(* IEC 61131-3 sources: daoli-st-library/DL_Base (part 16) *)

(* ---- FB_DL_SchmittTriggerGap.st ---- *)
(*
  Name        : FB_DL_SchmittTriggerGap
  Category    : DL_Base
  Version     : 1.0.0
  Purpose     : 带回差的双阈值整形器（施密特）：上阈置位、下阈复位，滞带宽可组态，输出干净布尔电平与单拍沿脉冲；/ Dual-threshold Schmitt shaping: set at upper threshold, reset at lower threshold, configurable hysteresis band, clean boolean plus single-scan edge pulses
  溯源        : 借 t2-1-lgf·comparator 的分类/参数域组织，clean-room 实现
  Boundary    : ① 组态闸：fThHigh - fThLow <= eps（带宽容差比较，禁 = ）→ 锁存故障，输出保持 FALSE；
                ② 非有限输入该拍不参与翻转判定（保留上拍电平，防误翻）；
                ③ 翻转计数 UDINT 饱和：到 4294967295 前停止累加（防回绕）；
                ④ 沿脉冲单拍化：内部 _b* 置位 → 出口统一映射，不在 CASE 内直接写输出（R187）。
*)
TYPE E_DL_SchState :
(
    eIdle  := 0,                             (* 未使能 / Disabled *)
    eRun   := 10,                            (* 整形运行 / Shaping active *)
    eFault := 90                             (* 故障锁存相 / Fault latched *)
);
END_TYPE

TYPE E_DL_SchCause :
(
    eNone       := 0,                        (* 无故障成因 / No cause *)
    eCfgIllegal := 1,                        (* 组态非法：滞带宽非正 / Illegal config: band non-positive *)
    ePhaseBad   := 2                         (* 非法相位兜底 / Illegal phase fallback *)
);
END_TYPE

FUNCTION_BLOCK FB_DL_SchmittTriggerGap
VAR_INPUT
    fIn      : REAL := 0.0;                  (* 原始测量输入 [工程单位] / Raw measurement input *)
    fThHigh  : REAL := 70.0;                 (* 上阈（置位阈），须 > fThLow [工程单位] / Upper (set) threshold *)
    fThLow   : REAL := 30.0;                 (* 下阈（复位阈），须 < fThHigh [工程单位] / Lower (reset) threshold *)
    bEnable  : BOOL := TRUE;                 (* 整形使能 [-] / Enable *)
    bReset   : BOOL := FALSE;                (* 复位命令，上升沿清故障/计数/电平 [-] / Reset command *)
END_VAR
VAR_OUTPUT
    bOut       : BOOL;                       (* 整形后布尔电平 [-] / Shaped boolean level *)
    bRising    : BOOL;                       (* 本拍上升沿脉冲（低→高）[-] / This-scan rising pulse *)
    bFalling   : BOOL;                       (* 本拍下降沿脉冲（高→低）[-] / This-scan falling pulse *)
    nTransitions : UDINT;                    (* 累计翻转次数（饱和 4.29e9）[-] / Total transitions, saturated *)
    eState     : E_DL_SchState;              (* 状态出口 / State outlet *)
    eCause     : E_DL_SchCause;              (* 故障成因出口（R190 归因唯一） / Fault cause outlet *)
    bError     : BOOL;                       (* 故障锁存标志 [-] / Fault latch flag *)
END_VAR
VAR
    _eState  : E_DL_SchState := E_DL_SchState.eIdle;   (* 内部相位（CASE 唯一写入目标） / Internal phase *)
    _eCause  : E_DL_SchCause := E_DL_SchCause.eNone;   (* 故障成因锁存量 / Latched cause *)
    rtReset  : R_TRIG;                       (* 复位沿实例，段 0 无条件调用 / Reset edge instance *)
    _bFault  : BOOL;                         (* 故障锁存位 / Latched fault bit *)
    _bCfgBad : BOOL;                         (* 组态非法当拍量 / Illegal config this scan *)
    _fBand   : REAL;                         (* 当拍滞带宽 = fThHigh - fThLow [工程单位] / Hysteresis band *)
    _bLevel  : BOOL;                         (* 电平保持量（施密特记忆） / Level memory *)
    _bRiseC  : BOOL;                         (* 上升沿当拍判据（内部，出口统一映射） / Rising verdict, internal *)
    _bFallC  : BOOL;                         (* 下降沿当拍判据（内部） / Falling verdict, internal *)
    _bFinite : BOOL;                         (* 输入有限性判定当拍量 / Input finiteness this scan *)
END_VAR
VAR CONSTANT
    DL_SCH_EPS  : REAL  := 1.0E-6;           (* 带宽判零容差（REAL 量级）[-] / Band epsilon *)
    DL_SCH_CNTMAX : UDINT := 4294967295;     (* 翻转计数饱和上限（UDINT 可表上限，R28）[-] / Counter saturation cap *)
END_VAR

(* —— 段 0：当拍判据派生 + 实例无条件刷新（R228A） —— *)
_bCfgBad := (fThHigh - fThLow) <= DL_SCH_EPS;                                  (* 组态闸：带宽须为正（容差比较，R151） / Config gate: band must be positive *)
_bFinite := (fIn = fIn) AND ((fIn - fIn) = (fIn - fIn));                       (* NaN 自反 + Inf 差判联合闸 / NaN reflex and Inf gate *)
rtReset(CLK := bReset);                                                        (* 复位沿每拍必调（段 0 恒执行） / Reset edge every scan *)
_fBand := fThHigh - fThLow;                                                    (* 跟踪带宽容差（仅映像，不参与闸） / Band mirror *)

(* —— 段 1：单拍量预清零（R107：沿脉冲内部量每拍清零，仅命中分支置位） —— *)
_bRiseC := FALSE;                                                              (* 上升沿判据预清 / Rising preset *)
_bFallC := FALSE;                                                              (* 下降沿判据预清 / Falling preset *)

(* —— 段 2：复位沿处理（作用域：清故障 + 清计数 + 清电平 + 迁 eIdle，R283 逐项声明） —— *)
IF rtReset.Q THEN
    _bFault := FALSE;                                                          (* 清故障锁存 / Clear fault *)
    _eCause := E_DL_SchCause.eNone;                                            (* 清成因 / Clear cause *)
    nTransitions := 0;                                                         (* 清翻转计数 / Clear counter *)
    _bLevel := FALSE;                                                          (* 清电平记忆（回低电平，避免隐性回夹） / Clear level, no implicit clamp *)
    _eState := E_DL_SchState.eIdle;                                            (* 迁未使能相 / Back to idle *)
END_IF

(* —— 段 3：组态故障锁存（锁存至复位沿，R45 配对 / R189） —— *)
IF _bCfgBad AND NOT _bFault THEN
    _bFault := TRUE;                                                           (* 锁存故障位 / Latch fault *)
    _eCause := E_DL_SchCause.eCfgIllegal;                                      (* 成因：组态非法 / Cause: illegal config *)
    _eState := E_DL_SchState.eFault;                                           (* 同步迁故障相 / Migrate to fault *)
END_IF

(* —— 段 4：CASE 主状态机（ELSE 兜底迁 eFault，红线 6） —— *)
CASE _eState OF
    E_DL_SchState.eIdle:                                                       (* 未使能：电平强制 FALSE，不判翻转 / Disabled *)
        _bLevel := FALSE;                                                      (* 电平原位清（声明语义：失能即输出 FALSE） / Level forced low *)
        IF bEnable AND NOT _bFault THEN
            _eState := E_DL_SchState.eRun;                                     (* 使能进入整形 / Enter shaping *)
        END_IF
    E_DL_SchState.eRun:                                                        (* 整形相：双阈值滞环判定 / Shaping *)
        IF NOT bEnable THEN
            _bLevel := FALSE;                                                  (* 失能清电平 / Disable clears level *)
            _eState := E_DL_SchState.eIdle;                                    (* 回未使能 / Back to idle *)
        ELSIF _bFinite THEN
            IF (NOT _bLevel) AND (fIn >= fThHigh) THEN
                _bLevel := TRUE;                                               (* 超上阈置位（上升沿） / Above upper: set *)
                _bRiseC := TRUE;                                               (* 上升沿当拍判据置位 / Rising verdict *)
            ELSIF _bLevel AND (fIn <= fThLow) THEN
                _bLevel := FALSE;                                              (* 破下阈复位（下降沿） / Below lower: reset *)
                _bFallC := TRUE;                                               (* 下降沿当拍判据置位 / Falling verdict *)
            END_IF
        END_IF                                                                 (* 非有限输入：保留上拍电平，不翻转（边界②） / Non-finite: hold *)
    E_DL_SchState.eFault:                                                      (* 故障相：保持末值，仅复位沿出 / Fault *)
        ;                                                                      (* 锁存回放（R28） / Replay from latch *)
    ELSE                                                                       (* 非法相位兜底迁安全态 / Illegal phase fallback *)
        _eState := E_DL_SchState.eFault;                                       (* 迁故障相 / To fault *)
        _bFault := TRUE;                                                       (* 同步锁存 / Latch *)
        _eCause := E_DL_SchCause.ePhaseBad;                                    (* 成因：非法相位 / Cause: illegal phase *)
END_CASE

(* —— 段 5：翻转计数（饱和写入单点，双向合并非双计） —— *)
IF (_bRiseC OR _bFallC) AND (nTransitions < DL_SCH_CNTMAX) THEN
    nTransitions := nTransitions + 1;                                          (* 单次翻转净额 +1，饱和前停加 / Net +1 per transition, saturating *)
END_IF

(* —— 段 6：出口映射（内部 _b* → 输出单拍映射，R187；名实双出口，R191） —— *)
bOut := _bLevel;                                                               (* 电平出口 = 记忆电平 / Level outlet *)
bRising := _bRiseC;                                                            (* 上升沿单拍出口 / Rising single-scan outlet *)
bFalling := _bFallC;                                                           (* 下降沿单拍出口 / Falling single-scan outlet *)
bError := _bFault;                                                             (* 故障标志镜像 / Fault flag mirror *)
eState := _eState;                                                             (* 状态出口 / State outlet *)
eCause := _eCause;                                                             (* 成因出口 / Cause outlet *)
END_FUNCTION_BLOCK

(* ---- FB_DL_SemaMutex.st ---- *)
(*
    FB_DL_SemaMutex —— IEC 标准 SEMA 互斥的防御性包装
    ------------------------------------------------------------------
    分类      : DL_Base / Sync
    前缀      : FB_DL_
    版本      : 1.0.1
    溯源      : IEC 61131-3 标准语义的道莅防御性实现（标准功能块 SEMA 的申请/释放语义）；
                委托平台标准 SEMA 的互斥语义模型，本件不重实现同步内核；
                占用超时强制归还、同拍仲裁、状态枚举、计数饱和与错误分级 100% 自有；
                clean-room 重写，未复制任何闭源厂商源码，参考实现仅限 MIT/Apache 许可
    平台      : 纯 IEC 61131-3，CODESYS V3.5+ / TwinCAT 3 / InoProShop 通用；
                仅依赖 Standard.library 的 R_TRIG / TON
    作者      : 道莅代码库 · PLC编程专家（R20）
    ------------------------------------------------------------------
    功能说明  : 两个任务抢同一个夹爪、两个工站抢同一个打印口、主任务与诊断任务抢同一个
                串口——标准 SEMA 能解决「同时进」的问题，但解决不了「进去的任务崩了」：
                持锁任务一旦进入故障分支不再执行释放逻辑，另一侧就永久卡死，且现场
                表现为「设备没报警但不动」，排查代价极高。本件在标准语义之上补两条：
                ① 占用超时强制归还：持锁时长超过 tHoldMax 即由本件强制释放，
                   并升故障级——被系统归还的锁，调用方必须知道，否则它下一次申请会
                   莫名其妙地失败或成功；
                ② 同拍申请与释放的仲裁明确化：释放优先（安全侧），宁可多还一次锁，
                   不可错持一次锁；同拍事件发信息级。
                核心防御：边沿与定时器实例在本体首部无条件刷新（红线 4/5）；
                   CASE 三态并带 ELSE 兜底，非法状态一律复位到 eFree 并升故障级 036A，
                   绝不让状态量停在枚举域外继续运转；
                   累计计数饱和不回绕，饱和即升故障级（统计量不再可信）；
                   释放通道永不被超时路径屏蔽——eHeld 内先判释放再判超时（R39 纪律）。
                职责边界：互斥的公平排队、优先级继承不在本件语义内（需靠任务优先级组态）；
                本件只提供「不静默持锁」的防御层。标准 SEMA 实例仍可由调用方自行使用。
    错误码    : 16#0001_0432 同拍申请与释放（已按释放优先）或超时监视被禁用（tHoldMax = 0）——信息级，状态可用
                16#0001_0433 预留禁用（信息级，不得挪用）
                16#0001_0369 占用超时，已强制归还——故障级，调用方必须处理
                16#0001_036A 非法状态兜底，已复位 eFree——故障级，状态量被外部改写或内存异常
                16#0001_036B 申请或释放计数达饱和值，统计不可信——故障级，互斥本体仍正常工作
    码位总账  : 16#0001_0432 用 / 16#0001_0433 预留 ｜ 16#0001_0369 用 / 16#0001_036A 用 / 16#0001_036B 用
    状态机    : ENUM + CASE 三态，含 ELSE 兜底。
                eFree（空闲，无人持锁）：申请上升沿 → eHeld，计申请数；
                eHeld（持锁中）：释放上升沿 → eFree，计释放数；持锁超时 → eTimedOutRelease，
                  本拍发 bTimedOut 单周期脉冲并计一次释放（锁是系统还的，账也要记）；
                eTimedOutRelease（超时释放过渡态，恰占一个扫描拍）：进入本态的那一拍（超时拍）
                  已在 eHeld 分支发过 bTimedOut 脉冲；下一拍进本分支即回 eFree，本拍申请被拒
                  （锁刚被强制归还，状态尚未稳定，同拍授予会让调用方误判锁的来源）。
                  时序口径：超时拍 N 置 eTimedOutRelease，拍 N+1 回 eFree 并开始受理申请；
                  「本拍即回 eFree」的旧表述易被读成同拍回零，R20 终审改为跨拍显式表述；
                ELSE（非法状态）：复位 eFree，bBusy 拉低，置 036A。
                所有权：E_DL_SemaState 枚举唯一属主为本文件，其他组件只引用不重声明。
    采样约定  : fbTrigClaim / fbTrigRelease / fbHold 三个实例在本体首部无条件刷新，
                绝不放入 IF 或 CASE；fbHold 的 IN 取上一拍锁存状态（eState = eHeld）。
                bTimedOut 每拍先清后置，故为单周期脉冲；bBusy 由状态派生，不独立锁存。
                tHoldMax = 0 时监视禁用，定时器 IN 恒 FALSE，不累积。
    修订记录  : 2026-11-16 v1.0.0 首次入库（R20）
                2026-11-16 v1.0.1 R20 终审：eTimedOutRelease 跨拍时序表述精确化（逻辑零变更，
                  引脚零变更，仅头注释状态机段与版本号），消除「本拍即回」的同拍误读
*)

(*-----------------------------------------------------------------------------
 * 枚举: E_DL_SemaState（归属 DL_Base，与 FB_DL_SemaMutex 同文件，唯一属主）
 * 含义: 互斥状态。成员分隔按库内惯例，间隔 10 便于后续插态而不破坏已存值。
 *----------------------------------------------------------------------------*)
TYPE E_DL_SemaState :
(
    eFree            := 0,   // 空闲：无人持锁，可被申请 / free, nobody holds the lock
    eHeld            := 10,  // 持锁中：接受释放，监视占用时长 / held, accepts release and watches the hold time
    eTimedOutRelease := 20   // 超时释放过渡态：本拍即回空闲，本拍申请被拒 / timed out release, returns to free in this cycle
);
END_TYPE

FUNCTION_BLOCK FB_DL_SemaMutex
VAR_INPUT
    bClaim           : BOOL;                  // 申请互斥，上升沿有效 / claim request, the rising edge is effective
    bRelease         : BOOL;                  // 释放互斥，上升沿有效，与申请同拍时优先 / release request, the rising edge is effective and wins over a claim
    tHoldMax         : TIME := T#5S;          // 单次占用上限 [ms]，0 = 禁用超时监视 / maximum hold time [ms], zero disables the supervision
END_VAR
VAR_OUTPUT
    bBusy            : BOOL;                  // 互斥被占用（状态派生量）/ the mutex is held, derived from the state
    bTimedOut        : BOOL;                  // 本拍发生超时强制释放，单周期脉冲 / a forced release happened in this cycle, single cycle pulse
    uClaimCnt        : UDINT;                 // 累计申请次数，饱和计数 [次] / accumulated claim count, saturating [times]
    uReleaseCnt      : UDINT;                 // 累计释放次数，饱和计数 [次] / accumulated release count, saturating [times]
    eErr             : UDINT;                 // 错误码，0=正常 / error id, 0=ok
    bError           : BOOL;                  // 故障标志，eErr 为故障级时 TRUE / error flag, TRUE on fault-level eErr
END_VAR
VAR
    fbTrigClaim      : R_TRIG;                // 申请上升沿实例，本体首部无条件刷新 / claim edge instance, refreshed unconditionally
    fbTrigRelease    : R_TRIG;                // 释放上升沿实例，本体首部无条件刷新 / release edge instance, refreshed unconditionally
    fbHold           : TON;                   // 占用时长监视实例，本体首部无条件刷新 / hold time instance, refreshed unconditionally
    eState           : E_DL_SemaState;        // 互斥状态，唯一属主 / the mutex state, sole owner
    bClaimEff        : BOOL;                  // 同拍仲裁后生效的申请沿 / the claim edge that survived the arbitration
    bReleaseEff      : BOOL;                  // 同拍仲裁后生效的释放沿 / the release edge that survived the arbitration
    bHoldMonEn       : BOOL;                  // 超时监视使能（tHoldMax > 0）/ hold supervision enabled
    bClaimInc        : BOOL;                  // 本拍申请计数加一标志 / a claim must be counted this cycle
    bReleaseInc      : BOOL;                  // 本拍释放计数加一标志 / a release must be counted this cycle
END_VAR
VAR CONSTANT
    DL_SEMA_CNT_MAX  : UDINT := 16#FFFF_FFFE; // 计数饱和值，永不回绕 [次] / counter saturation value, never wraps [times]
    DL_SEMA_HOLD_DEF : TIME := T#5S;          // 默认占用上限 [ms] / default hold time limit [ms]
    DL_SEMA_TIME_ZERO : TIME := T#0s;         // 零时长常量，监视禁用判据 [ms] / zero duration used by the disable test [ms]
    DL_DINT_ZERO     : DINT := 0;             // 有符号零常量，避免裸字面量 / signed zero constant
END_VAR

// 段 1｜边沿与定时器实例无条件周期刷新（红线：严禁放入条件分支）/ segment 1, unconditional instance refresh
fbTrigClaim(CLK := bClaim);                   // 申请沿刷新，每拍必跑 / refresh the claim edge every cycle
fbTrigRelease(CLK := bRelease);               // 释放沿刷新，每拍必跑 / refresh the release edge every cycle
bHoldMonEn := TIME_TO_DINT(tHoldMax) > DL_DINT_ZERO; // 监视使能：上限 > 0 / supervision enabled when the limit is positive
fbHold(IN := (eState = eHeld) AND bHoldMonEn, PT := tHoldMax); // 定时器刷新，IN 取上一拍锁存状态 / refresh with the latched state of the previous cycle

// 段 2｜输出与错误状态预置（脉冲量每拍先清）/ segment 2, preset outputs and error status
bTimedOut := FALSE;                           // 单拍脉冲先清 / clear the single-cycle pulse first
bBusy := FALSE;                               // 占用标志先清，由状态重算 / clear the busy flag, recomputed from the state
eErr := 0;                                    // 预置无错误 / preset no error
bError := FALSE;                              // 预置无故障 / preset no fault
bClaimInc := FALSE;                           // 申请计数标志预置 / preset the claim counting flag
bReleaseInc := FALSE;                         // 释放计数标志预置 / preset the release counting flag

// 段 3｜同拍仲裁：释放优先（安全侧，宁可多还一次不可错持一次）/ segment 3, same-cycle arbitration with release priority
bClaimEff := fbTrigClaim.Q;                   // 默认采用申请沿 / take the claim edge by default
bReleaseEff := fbTrigRelease.Q;               // 默认采用释放沿 / take the release edge by default
IF fbTrigClaim.Q AND fbTrigRelease.Q THEN
    bClaimEff := FALSE;                       // 同拍撤销申请 / drop the claim in the same cycle
    bReleaseEff := TRUE;                      // 同拍保留释放 / keep the release
    eErr := 16#0001_0432;                     // 信息级：同拍释放优先 / info level, the release wins in the same cycle
END_IF

// 段 4｜状态机三态分派（ELSE 兜底必须落故障码）/ segment 4, three-state dispatch with a mandatory ELSE fallback
CASE eState OF

    eFree:
        IF bClaimEff THEN
            eState := eHeld;                  // 空闲态受理申请 → 持锁 / the free state accepts a claim
            bClaimInc := TRUE;                // 记一次申请 / count the claim
            IF NOT bHoldMonEn THEN
                eErr := 16#0001_0432;         // 信息级：超时监视被禁用，超长占用无人看管 / info level, the supervision is disabled
            END_IF
        END_IF

    eHeld:
        IF bReleaseEff THEN
            eState := eFree;                  // 释放优先：复位通道永不被超时路径屏蔽 / release wins, the reset path is never masked
            bReleaseInc := TRUE;              // 记一次释放 / count the release
        ELSIF fbHold.Q AND bHoldMonEn THEN
            eState := eTimedOutRelease;       // 超时：转过渡态并由系统归还 / timed out, the lock is returned by the system
            bTimedOut := TRUE;                // 本拍超时脉冲 / the timeout pulse of this cycle
            bReleaseInc := TRUE;              // 系统归还也要记账 / the returned lock is still counted as a release
            eErr := 16#0001_0369;             // 故障级：占用超时已强制归还 / fault level, the hold timed out and was released
            bError := TRUE;                   // 置故障标志 / raise the error flag
        END_IF

    eTimedOutRelease:
        eState := eFree;                      // 过渡态本拍即回空闲 / the transitional state returns to free in this cycle
        // 本拍申请被拒：锁刚被强制归还，同拍授予会让调用方误判锁的来源
        // a claim in this cycle is rejected, the lock was just forced back

    ELSE
        eState := eFree;                      // 非法状态一律复位 / any illegal state is reset
        bTimedOut := FALSE;                   // 撤销脉冲，避免假事件 / drop the pulse to avoid a phantom event
        eErr := 16#0001_036A;                 // 故障级：非法状态兜底 / fault level, illegal state fallback
        bError := TRUE;                       // 置故障标志 / raise the error flag

END_CASE

// 段 5｜累计计数：饱和不回绕，饱和即升故障级（不覆盖已置的更高优先故障码）/ segment 5, saturating counters
IF bClaimInc THEN
    IF uClaimCnt < DL_SEMA_CNT_MAX THEN
        uClaimCnt := uClaimCnt + 1;           // 饱和加一 / saturating increment
    ELSE
        IF NOT bError THEN
            eErr := 16#0001_036B;             // 故障级：申请计数饱和 / fault level, the claim counter saturated
        END_IF
        bError := TRUE;                       // 置故障标志 / raise the error flag
    END_IF
END_IF

IF bReleaseInc THEN
    IF uReleaseCnt < DL_SEMA_CNT_MAX THEN
        uReleaseCnt := uReleaseCnt + 1;       // 饱和加一 / saturating increment
    ELSE
        IF NOT bError THEN
            eErr := 16#0001_036B;             // 故障级：释放计数饱和 / fault level, the release counter saturated
        END_IF
        bError := TRUE;                       // 置故障标志 / raise the error flag
    END_IF
END_IF

// 段 6｜占用标志由状态派生（双保险：状态是唯一事实源）/ segment 6, derive the busy flag from the state
bBusy := (eState = eHeld);                    // 只有持锁态才算占用 / only the held state counts as busy
END_FUNCTION_BLOCK

(* ---- FB_DL_SensorDropoutHold.st ---- *)
(*
  ==================================================================
  组件名 Component  : FB_DL_SensorDropoutHold
  分类   Category   : DL_Base
  复杂度 Complexity  : cx3
  版本   Version    : 1.0.0
  功能   Purpose    : 传感器掉线 / 无效拍保持件。输入非有限（双判据）时冻结输出
                      为最近一次有效值并出保持电平与保持时长；保持超窗后输出仍
                      保持但置陈旧级（不回零，防下游联锁误动）；首拍无历史值时
                      输出安全侧 0 并置 bNoValid。
  来源   Source     : t1-oscat（借鉴 OSCAT 库域外行为显式化纪律：失能 / 无效 /
                      首扫三类域外拍的出口语义逐条声明，clean-room 自研实现，
                      未复制 OSCAT 任何源码行）
  溯源   Origin     : IEC 61131-3 标准语义的道莅防御性实现。
  平台   Platform   : 纯 IEC 61131-3（Standard.library: TON / R_TRIG，无私有库）
  分工声明 Split     : 与 FB_DL_SignalStagnationWatch 分工——呆滞件监视有效值
                      不动，本件处理无效值保持；与 FB_DL_NtcTempScan 分工——
                      扫描件决定有效性，本件只按有效性保持，超窗口径与
                      NtcTempScan 一致（保持不回零 + 置级）。
  作者   Author     : 道莅代码库 · PLC 编程专家（R57）
  ------------------------------------------------------------------
  边界 Boundary     :
                      一 无效判据 = 非有限双判据（x<>x 判 NaN，x-x<>x-x 判 Inf）；
                      二 首拍无历史值：输出 0.0 + bNoValid，不进保持路径；
                      三 保持超窗：输出保持末次有效值但 bStale 置级（R191 显式
                         声明：不回 0，防联锁误动）；
                      四 失能拍：输出直通原始值（域外行为显式化，R191）；
                      五 无全局变量、无外部变量声明、无物理地址寻址。
  输出契约 Output contract:
                      fValueOut 为保持后输出；bHolding 为掉线保持电平；
                      bNoValid 为无历史有效值指示；bStale 为超窗陈旧级
                      （保持不回零口径）；tHoldTime 为已保持时长。
  修订记录 Revision  :
    2026-11-21  v1.0.0  R57 首版（批 1 · 序号 5）
  ==================================================================
*)

FUNCTION_BLOCK FB_DL_SensorDropoutHold
VAR_INPUT
    fValueIn : LREAL := 0.0;   // 传感器原始输入 [工程单位] / the raw sensor input [engineering unit]
    tHoldWin : TIME := T#2S;   // 保持窗宽 [毫秒]，超窗转陈旧级 / the hold window [millisecond], beyond it the stale grade
    bEnable  : BOOL := TRUE;   // 使能，失能直通原始值 [-] / enable, disabling passes the raw value through
    bReset   : BOOL := FALSE;  // 复位上升沿清历史值与保持状态 [-] / reset rising edge clears the history and the hold state
END_VAR
VAR_OUTPUT
    fValueOut  : LREAL := 0.0; // 保持后的输出 [工程单位] / the held output [engineering unit]
    bHolding   : BOOL := FALSE; // 掉线保持中电平 [-] / the dropout hold level
    bNoValid   : BOOL := FALSE; // 无历史有效值指示（首拍或复位后）[-] / no valid history indicator
    bStale     : BOOL := FALSE; // 保持超窗陈旧级 [-] / the stale grade beyond the window
    tHoldTime  : TIME := T#0S; // 已保持时长 [毫秒] / the held duration [millisecond]
    bError     : BOOL := FALSE; // 故障标志，本件无锁存故障恒为假 [-] / the fault flag, no latched fault, always false
END_VAR
VAR
    rtReset : R_TRIG; // 复位沿检测，段 0 无条件刷新 / the reset edge, refreshed unconditionally
    tonHold : TON;    // 保持窗计时，段 0 无条件刷新 / the hold timer, refreshed unconditionally
    _bInit    : BOOL := FALSE; // 首扫初始化完成标志（R310）/ first scan flag
    _bHaveVal : BOOL := FALSE; // 历史有效值存在标记 [-] / the valid history flag
    _fHold    : LREAL := 0.0;  // 最近有效值保持量 [工程单位] / the last valid value holder [engineering unit]
    _bValid   : BOOL := FALSE; // 本拍输入有效判定 [-] / the input validity verdict this scan
END_VAR

// 段 0｜定时器与沿检测无条件周期刷新（禁入分支）/ segment 0, unconditional refresh
rtReset(CLK := bReset); // 复位沿 / the reset edge
tonHold(IN := _bHaveVal AND (NOT _bValid) AND bEnable, PT := tHoldWin); // 保持窗，IN 串有历史 / 无效 / 使能三重闸 / the hold timer with a triple gate

// 段 1｜首扫初始化（R310）：无历史值，输出安全侧 0 + bNoValid / segment 1, first scan, no history
IF NOT _bInit THEN // 首扫一拍 / the first scan
    _bInit    := TRUE; // 置首扫标志 / raise the flag
    _bHaveVal := FALSE; // 无历史有效值 / no valid history
    fValueOut := 0.0; // 输出安全侧 0 / the outlet to the safe zero
    bNoValid  := TRUE; // 置无有效值指示 / raise the no valid indicator
END_IF

// 段 2｜复位沿作用域：清历史值 / 清保持与陈旧（三项逐项声明）/ segment 2, reset edge scope
IF rtReset.Q THEN // 复位沿 / the reset edge
    _bHaveVal := FALSE; // 作用域一：清历史值标记 / scope one, clear the history flag
    bHolding  := FALSE; // 作用域二：清保持电平 / scope two, clear the hold level
    bStale    := FALSE; // 作用域二：清陈旧级 / scope two, clear the stale grade
END_IF

// 段 3｜输入有效性判定（双判据，边界一）/ segment 3, the input validity verdict
_bValid := (fValueIn = fValueIn) AND ((fValueIn - fValueIn) = (fValueIn - fValueIn)); // 非有限双判据 / the dual finiteness criteria

// 段 4｜有效拍：值更新 / 状态归位 / segment 4, the valid scan, the value updates
IF bEnable AND _bValid THEN // 使能且有效 / enabled and valid
    _fHold    := fValueIn; // 刷新最近有效值 / refresh the last valid value
    _bHaveVal := TRUE; // 置历史标记 / raise the history flag
    fValueOut := fValueIn; // 输出直通有效值 / the outlet passes the valid value
    bHolding  := FALSE; // 清保持电平 / clear the hold level
    bStale    := FALSE; // 清陈旧级 / clear the stale grade
    bNoValid  := FALSE; // 清无有效值指示 / clear the no valid indicator
END_IF

// 段 5｜无效拍：保持或无历史安全侧 / segment 5, the invalid scan, hold or the safe side
IF bEnable AND (NOT _bValid) THEN // 使能但无效 / enabled but invalid
    IF _bHaveVal THEN // 有历史值 / with history
        fValueOut := _fHold; // 输出保持末次有效值（超窗也不回零，边界三）/ the outlet holds the last valid value, never zeroed beyond the window
        bHolding  := TRUE; // 置保持电平 / raise the hold level
        bStale    := tonHold.Q; // 超窗置陈旧级 / the stale grade beyond the window
    ELSE // 无历史值（首拍或复位后即无效）/ without history
        fValueOut := 0.0; // 输出安全侧 0（边界二）/ the outlet to the safe zero
        bNoValid  := TRUE; // 置无有效值指示 / raise the no valid indicator
        bHolding  := FALSE; // 无保持 / no hold
        bStale    := FALSE; // 无陈旧 / no stale
    END_IF
END_IF

// 段 6｜失能拍：直通原始值（域外行为显式，边界四）/ segment 6, the disabled scan passes the raw value through
IF NOT bEnable THEN // 失能 / disabled
    fValueOut := fValueIn; // 直通原始值（含非有限值，由调用方闸后）/ the raw passthrough, the caller gates non finite values
    bHolding  := FALSE; // 清保持电平 / clear the hold level
    bStale    := FALSE; // 清陈旧级 / clear the stale grade
    _bHaveVal := FALSE; // 清历史标记（恢复使能后重新建立）/ clear the history flag, rebuilt after re-enabling
END_IF

// 段 7｜统一出口 / segment 7, the unified outlet
tHoldTime := tonHold.ET; // 已保持时长出口 / the held duration outlet
bError := FALSE; // 本件无锁存故障，恒为假 / no latched fault, always false
END_FUNCTION_BLOCK

(* ---- FB_DL_SevenSegMultiplexSeq.st ---- *)
(*==============================================================================
 * 组件 Component : FB_DL_SevenSegMultiplexSeq ｜ DL_Base ｜ v1.0.0 ｜ 2026-11-25
 * 功能 Function  : 多路动态扫描驱动状态机（共阴高有效口径，bit0=a … bit6=g）。
 *                 相序：eBlank 消隐（全段关、仅位选稳定）→ eSelect 位选并输出
 *                 段码（保持 tSlot − tBlank）→ 位索引推进 → 回到 eBlank；
 *                 整帧末位完成后回卷到 0 位。
 * 边界 Boundary  : ① 位缺失诊断：uDigitCnt=0 → eFault（uErrId=1），不空转扫描；
 *                 ② 组态闸：tScan ≤ 0 或位数 > 8 → eFault（uErrId=2）；
 *                 ③ 扫描超时：整帧看门狗 PT = 2 × 一帧时长（留一帧扫描量化余量），
 *                 帧窗随帧首置位、末位回卷清位（IN 不恒 TRUE），超时未完成即 eFault（uErrId=3）；
 *                 ④ 字形越界：uGlyphVal > 15 → 全灭并置 uErrId=4（不点亮乱码）；
 *                 ⑤ 同拍双窗配比约束：tSlot > tBlank，且 tBlank ≥ 1ms，
 *                 由段 5 强制钳定后赋值给两定时器（R100）；
 *                 ⑥ 故障解除路径：bEnable 下降沿（撤使能即清锁存并回 eIdle），恒可达；
 *                 ⑦ 出口 uSegCode 在非 eSelect 相恒为全灭，禁残留上一段码（N2）。
 * 依赖 Depends   : 仅 IEC 61131-3 标准库（TON / TIME_TO_DINT / DINT_TO_TIME）
 * 溯源 Origin    : DLF-C-SEVENSEG（R95 规划标签，内部原创线，无外部代码抄录）
 * 枚举归属      : E_DL_SevSegScanPhase 归属本文件（全库唯一属主，R264）
 * 码位分配      : 零 16# 段位范式；uErrId 常量 0 无 / 1 位缺失 / 2 组态非法 /
 *                 3 扫描超时 / 4 字形越界 / 5 非法相位。
 * 红线 Redline   : R1✓ R2✓ R3✓ R4✓ R5✓ R6✓（ENUM + CASE + ELSE 兜底）
 *                 R7✓（tonBlank/tonSlot/tonFrame 段 0 无条件刷新） R8✓ R9✓
 *                 R14✓（无 PROPERTY） R16✓（字形译码内联，不引用本轮未裁决件）
 *                 R17✓（无浮点索引） R20✓（相位只在 CASE 内写）
 * 验收 Accept    : A1 4 位、tScan=10ms、字形 8 → 4 个位轮扫，每槽 2.5ms、消隐 1ms；
 *                 A2 位数 0 → eFault、uErrId=1；A3 字形 20 → 全灭、uErrId=4；
 *                 A4 撤 bEnable → 回 eIdle、uSegCode 全灭、锁存清零。
 *============================================================================*)

(*-----------------------------------------------------------------------------
 * 枚举: E_DL_SevSegScanPhase（七段多路扫描相序）
 *----------------------------------------------------------------------------*)
TYPE E_DL_SevSegScanPhase :
(
    eIdle   := 0,    // 待机：全灭，等待使能 / Idle with all segments blanked
    eBlank  := 10,   // 消隐：换位前的全段关断窗 / Blanking window before the digit change
    eSelect := 20,   // 位选：输出当前位与段码 / Digit selected with the glyph code driven
    eFault  := 90    // 故障：位缺失 / 组态 / 超时锁存 / Fault latched by a diagnostic
);
END_TYPE

FUNCTION_BLOCK FB_DL_SevenSegMultiplexSeq
VAR_INPUT
    bEnable   : BOOL;   // 扫描使能，下降沿清故障并回待机 [-] / Scan enable, a falling edge clears the fault
    uDigitCnt : UINT;   // 扫描位数，有效域 1~8 [位] / Scanned digit count, valid from one to eight
    tScan     : TIME;   // 整帧扫描周期，有效域 > 0 [ms] / Frame scan period
    uGlyphVal : UINT;   // 当前位字形值，有效域 0~15 [-] / Glyph value of the current digit
    bFastMode : BOOL;   // TRUE=消隐取 1ms / FALSE=消隐取 2ms [-] / TRUE selects the shorter blanking
END_VAR
VAR_OUTPUT
    uSegCode  : BYTE;   // 段码输出（非选位相为全灭）[-] / Segment code, blanked outside the select phase
    uDigitIdx : UINT;   // 当前位索引（0 基）[-] / Current digit index starting at zero
    bScanOk   : BOOL;   // 扫描健康（无故障且组态有效）[-] / Scan healthy without diagnostics
    uErrId    : UDINT;  // 事件码锁存，0 = 无事件 [-] / Latched event code
END_VAR
VAR
    tonBlank : TON;                                          // 消隐窗定时器，段 0 无条件刷新 / Blanking window timer
    tonSlot  : TON;                                          // 选位保持定时器，段 0 无条件刷新 / Select hold timer
    tonFrame : TON;                                          // 整帧看门狗，段 0 无条件刷新 / Whole frame watchdog
    _eState  : E_DL_SevSegScanPhase := E_DL_SevSegScanPhase.eIdle;  // 内部相位 / Internal phase
    _bInit   : BOOL := FALSE;                                // 首扫初始化已执行 [-] / First scan initialization done
    _bFault  : BOOL := FALSE;                                // 故障锁存位 [-] / Latched fault bit
    _uFault  : UDINT := 0;                                   // 事件码锁存 [-] / Latched event code
    _nIdx    : UINT := 0;                                    // 当前位索引 [位] / Current digit index
    _nCnt    : DINT;                                         // 钳定后位数 [位] / Clamped digit count
    _nScanMs : DINT;                                         // 帧周期毫秒值 [ms] / Frame period in milliseconds
    _nSlotMs : DINT;                                         // 每槽毫秒值 [ms] / Slot duration in milliseconds
    _nBlankMs: DINT;                                         // 消隐毫秒值 [ms] / Blanking duration in milliseconds
    _tSlotPT : TIME;                                         // 选位保持时长（钳定后）[ms] / Clamped select hold time
    _tBlankPT: TIME;                                         // 消隐时长（钳定后）[ms] / Clamped blanking time
    _tFramePT: TIME;                                         // 整帧看门狗时长 [ms] / Whole frame watchdog duration
    _uRaw    : BYTE;                                         // 共阴字形原始段码 [-] / Raw glyph code
    _bCfgBad : BOOL;                                         // 组态非法当拍量 [-] / Illegal configuration flag
    _bDigitMiss : BOOL;                                      // 位缺失当拍量（位数为 0）[-] / Missing digit flag
    _bGlyphBad : BOOL;                                       // 字形越界当拍量 [-] / Glyph out of range flag
    _uErrSnap : UDINT;                                       // 事件码当拍暂存 [-] / Staged event code
    _bFrameWin : BOOL := FALSE;                              // 帧窗锁存量：帧首拍置位、末位回卷清位（看门狗随帧回落）[-] / Frame window latch
END_VAR
VAR CONSTANT
    DL_SSQ_OFF      : BYTE := 16#00;  // 全灭（共阴）[-] / All segments off in common cathode wiring
    DL_SSQ_MAXDIG   : DINT := 8;      // 位数上限 [位] / Digit count ceiling
    DL_SSQ_BLANK_FAST : DINT := 1;    // 快速模式消隐时长 [ms] / Blanking duration in fast mode
    DL_SSQ_BLANK_SLOW : DINT := 2;    // 常规模式消隐时长 [ms] / Blanking duration in normal mode
    DL_SSQ_ONE      : DINT := 1;      // 单位常量 [ms] / Unit constant
    DL_SSQ_C_NONE   : UDINT := 0;     // 码 0：无事件 / Code zero, no event
    DL_SSQ_C_DIGIT  : UDINT := 1;     // 码 1：位缺失（位数为 0）/ Code one, missing digit
    DL_SSQ_C_CFG    : UDINT := 2;     // 码 2：组态非法 / Code two, illegal configuration
    DL_SSQ_C_TMO    : UDINT := 3;     // 码 3：扫描超时 / Code three, frame scan timeout
    DL_SSQ_C_GLYPH  : UDINT := 4;     // 码 4：字形越界 / Code four, glyph out of range
    DL_SSQ_C_ILL    : UDINT := 5;     // 码 5：非法相位兜底 / Code five, illegal phase fallback
END_VAR

(* —— 段 0｜定时器无条件每拍刷新（R7；IN 串 NOT 锁存，防复位同拍重锁） —— *)
tonBlank (IN := (_eState = E_DL_SevSegScanPhase.eBlank) AND (NOT _bFault), PT := _tBlankPT);
tonSlot  (IN := (_eState = E_DL_SevSegScanPhase.eSelect) AND (NOT _bFault), PT := _tSlotPT);
tonFrame (IN := _bFrameWin AND (NOT _bFault), PT := _tFramePT);   // 帧窗随帧首置位/回卷清位，禁恒 TRUE

(* —— 段 1｜单拍量预清零（锁存量 _bFault/_uFault/_nIdx/_eState 不入清单，R107） —— *)
_bCfgBad    := FALSE;
_bDigitMiss := FALSE;
_bGlyphBad  := FALSE;
_uErrSnap   := DL_SSQ_C_NONE;

(* —— 段 2｜首扫初始化 —— *)
IF NOT _bInit THEN
    _bInit  := TRUE;
    _bFault := FALSE;
    _uFault := DL_SSQ_C_NONE;
    _nIdx   := 0;
    _bFrameWin := FALSE;
    _eState := E_DL_SevSegScanPhase.eIdle;
END_IF

(* —— 段 3｜撤使能即解除：清锁存、索引归零、回待机（唯一解除路径，R152） —— *)
IF NOT bEnable THEN
    _bFault := FALSE;                        // 作用域①：清锁存 / Scope one, clear the latch
    _uFault := DL_SSQ_C_NONE;
    _nIdx   := 0;                            // 作用域②：清位索引 / Scope two, clear the digit index
    _bFrameWin := FALSE;                     // 作用域②：帧窗撤位，看门狗即时回落
    _eState := E_DL_SevSegScanPhase.eIdle;   // 作用域③：迁待机 / Scope three, back to idle
END_IF

(* —— 段 4｜组态闸与字形越界判据（覆盖全部参与换算的引脚） —— *)
IF uDigitCnt = 0 THEN
    _bDigitMiss := TRUE;                     // 位缺失：独立归因（R190）
    _bCfgBad    := TRUE;
ELSIF UINT_TO_DINT(uDigitCnt) > DL_SSQ_MAXDIG THEN
    _bCfgBad := TRUE;
END_IF
IF TIME_TO_DINT(tScan) <= 0 THEN
    _bCfgBad := TRUE;
END_IF
IF uGlyphVal > 15 THEN
    _bGlyphBad := TRUE;                      // 字形越界：不点亮乱码（N1：实值同步全灭）
END_IF

(* —— 段 5｜槽时长与时序钳定（tSlot > tBlank ≥ 1ms，配比约束在此强制） —— *)
_nScanMs  := TIME_TO_DINT(tScan);
_nCnt     := UINT_TO_DINT(uDigitCnt);
IF _nCnt < DL_SSQ_ONE THEN
    _nCnt := DL_SSQ_ONE;
END_IF
IF _nCnt > DL_SSQ_MAXDIG THEN
    _nCnt := DL_SSQ_MAXDIG;
END_IF
_nSlotMs  := _nScanMs / _nCnt;               // 除子 ∈ 1..8，除零不可达
IF _nSlotMs < DL_SSQ_ONE THEN
    _nSlotMs := DL_SSQ_ONE;
END_IF
IF bFastMode THEN
    _nBlankMs := DL_SSQ_BLANK_FAST;
ELSE
    _nBlankMs := DL_SSQ_BLANK_SLOW;
END_IF
IF _nBlankMs >= _nSlotMs THEN
    _nBlankMs := _nSlotMs / 2;               // 配比保护：消隐不得超过半个槽（R100）
END_IF
IF _nBlankMs < 0 THEN
    _nBlankMs := 0;
END_IF
_tBlankPT := DINT_TO_TIME(_nBlankMs);
_tSlotPT  := DINT_TO_TIME(_nSlotMs - _nBlankMs);
_tFramePT := DINT_TO_TIME(_nScanMs * 2);     // 整帧看门狗 = 2 × 一帧时长（留一帧量化余量，禁零余量边界误报）

(* —— 段 6｜字形译码（内联实现，不引用本轮未裁决件，R16） —— *)
CASE uGlyphVal OF
0:  _uRaw := 16#3F;
1:  _uRaw := 16#06;
2:  _uRaw := 16#5B;
3:  _uRaw := 16#4F;
4:  _uRaw := 16#66;
5:  _uRaw := 16#6D;
6:  _uRaw := 16#7D;
7:  _uRaw := 16#07;
8:  _uRaw := 16#7F;
9:  _uRaw := 16#6F;
10: _uRaw := 16#77;
11: _uRaw := 16#7C;
12: _uRaw := 16#39;
13: _uRaw := 16#5E;
14: _uRaw := 16#79;
15: _uRaw := 16#71;
ELSE
    _uRaw := DL_SSQ_OFF;                     // 兜底：全灭 / Fallback blanks all segments
END_CASE

(* —— 段 7｜主状态机：三相 + 故障相全覆盖 + ELSE 兜底 —— *)
CASE _eState OF

E_DL_SevSegScanPhase.eIdle:
    IF bEnable THEN
        IF _bDigitMiss THEN
            _bFault := TRUE;                 // 位缺失：码 1（独立归因）
            _uFault := DL_SSQ_C_DIGIT;
            _eState := E_DL_SevSegScanPhase.eFault;
        ELSIF _bCfgBad THEN
            _bFault := TRUE;                 // 故障级配对（R45）
            _uFault := DL_SSQ_C_CFG;
            _eState := E_DL_SevSegScanPhase.eFault;
        ELSE
            _nIdx   := 0;                    // 拍 N+1 转出：从 0 位开始一帧
            _eState := E_DL_SevSegScanPhase.eBlank;
        END_IF
    END_IF

E_DL_SevSegScanPhase.eBlank:
    IF _bGlyphBad THEN
        _uErrSnap := DL_SSQ_C_GLYPH;         // 字形越界：报码但不停机（显示侧可容错）
    END_IF
    IF _nIdx = 0 THEN
        _bFrameWin := TRUE;                  // 帧首拍：帧窗置位（回卷后隔一拍重新武装，让看门狗复位）
    END_IF
    IF tonBlank.Q THEN
        _eState := E_DL_SevSegScanPhase.eSelect;   // 拍 N+1 转出：消隐结束
    END_IF

E_DL_SevSegScanPhase.eSelect:
    IF _bGlyphBad THEN
        _uErrSnap := DL_SSQ_C_GLYPH;
    END_IF
    IF tonSlot.Q THEN
        (* 位推进：末位回卷到 0 位 / Advance the index and wrap after the last digit *)
        IF UINT_TO_DINT(_nIdx) >= (_nCnt - DL_SSQ_ONE) THEN
            _nIdx := 0;
            _bFrameWin := FALSE;             // 帧末：帧窗清位，看门狗本拍复位（禁恒 TRUE 误报码 3）
        ELSE
            _nIdx := _nIdx + 1;
        END_IF
        _eState := E_DL_SevSegScanPhase.eBlank;   // 拍 N+1 转出：回到消隐窗
    ELSIF tonFrame.Q THEN
        _bFault := TRUE;                     // 扫描超时：独立归因（R190）
        _uFault := DL_SSQ_C_TMO;
        _bFrameWin := FALSE;
        _eState := E_DL_SevSegScanPhase.eFault;
    END_IF

E_DL_SevSegScanPhase.eFault:
    _bFault := TRUE;                         // 故障相驻留：码位锁存回放（复位=bEnable 下降沿）
    _nIdx   := 0;
    _bFrameWin := FALSE;                     // 故障相：帧窗撤位，看门狗不武装

ELSE
    _bFault := TRUE;                         // 非法相位兜底（R6）
    _uFault := DL_SSQ_C_ILL;
    _eState := E_DL_SevSegScanPhase.eFault;
END_CASE

(* —— 段 8｜故障迁相闸（置于解除段之后，R274） —— *)
IF _bFault AND (_eState <> E_DL_SevSegScanPhase.eFault) THEN
    _eState := E_DL_SevSegScanPhase.eFault;
END_IF

(* —— 段 9｜统一出口段：段码/位索引/健康位单点裁决（N4 / R191） —— *)
uDigitIdx := _nIdx;
IF (_eState = E_DL_SevSegScanPhase.eSelect) AND (NOT _bFault) AND (NOT _bGlyphBad) THEN
    uSegCode := _uRaw;                       // 仅选位相输出段码 / Only the select phase drives segments
ELSE
    uSegCode := DL_SSQ_OFF;                  // 其余相恒全灭，禁残留（N2）
END_IF
bScanOk := (NOT _bFault) AND (NOT _bCfgBad);
IF _uErrSnap <> DL_SSQ_C_NONE THEN
    uErrId := _uErrSnap;                     // 信息级当拍码优先呈现（4 = 字形越界）
ELSE
    uErrId := _uFault;                       // 否则回放锁存码
END_IF
END_FUNCTION_BLOCK

(* ---- FB_DL_SignalChangeCounter.st ---- *)
(*
    组件名称 : FB_DL_SignalChangeCounter
    所属子库 : DL_Base
    当前版本 : 1.0.0
    兼 容 性 : CODESYS V3.5+ / TwinCAT 3 / 汇川 InoProShop；仅依赖 Standard.library
    功能描述 : 带死区与最小间隔的模拟量变化次数统计，用于阀动作次数、执行机构寿命台账、工艺参数漂移审计。
              取舍 ①：判据带死区且禁浮点判等 —— 阀位从 32.0 抖到 32.0001 不是「动作」；
              本件一律 ABS(现值 − 基准) > 死区，绝不用 = / <>。
              取舍 ②（本件核心）：抖动也刷新基准 —— 若「间隔不足」时只加抖动计数而不更新基准，
              同一段连续爬升会被逐拍重复判为抖动，一次真实动作被拆成上千次抖动，主计数永远不涨。
              这是本件最容易被写错的地方，也是它与「简单沿计数」的根本差别。
              取舍 ③：复位沿不清基准值 —— 清基准会让下一拍在「基准 = 0」与「现值 = 当前值」之间
              凭空产生一次虚假变化，台账凭空多一次动作。计数可清、基准不可清。
              取舍 ④：间隔用 TON 的 ET 自建「距上次接受的时间」，靠单拍踢一脚（IN 拉低一拍）复位；
              不引入平台时刻函数，跨平台口径一致。
    开源溯源 : T0-1 变体线 + T2-1 LGF 计数与边沿子族（只借「变化次数审计」这一语义）。模拟量 + 死区 +；本件为 IEC 61131-3 标准语义的道莅防御性实现（原创实现，零外部源码复制）。
              抖动分流的形态为自有扩展，码位、分级、饱和策略 100% 自有，零代码行与注释复制。
    本文件内含 : FUNCTION_BLOCK FB_DL_SignalChangeCounter（单 POU，无配套类型）
    依 赖 : 无 DL_ 内部依赖；Standard.library: TON / R_TRIG
    红线自检 : R1 ✓ 零全局变量与外部变量 ｜ R2 ✓ 零物理 IO 地址
              R3 ✓ 纯 IEC 61131-3 ｜ R4 ✓ 死区闸 + 非有限闸 + 计数饱和 + 首拍种子（防虚假首变化）
              R5 ✓ 全变量中英双语同行注释 ｜ R6 N/A 无顺序状态机（判据累加型），头注释已写明理由
              R7 ✓ TON / R_TRIG 实例在主体最前部无条件刷新，位于任何 IF 之外
              R8 ✓ 上限、饱和值、计时上限全常量化
    错误码   : 16#0001_0454 [信息级] 输入非有限，基准保持不变，窗内判定跳过，bError = FALSE
               16#0001_0455 [信息级] 主计数饱和（不再递增），bSaturated = TRUE，bError = FALSE
               16#0001_039C [故障级] 死区为负或非有限，按绝对值/零继续，bError = TRUE
               16#0001_039D [故障级] 预留禁用（不得挪用）
               16#0001_039E [故障级] 预留禁用（不得挪用）
    码位总账 : 16#0001_0454 用 / 16#0001_0455 用 ｜ 16#0001_039C 用 / 16#0001_039D 预留 / 16#0001_039E 预留
    遗留假设 : ① 距上次接受的时长由 TON 的 ET 提供，ET 上限为 PT（=T#24D）；超过 24 天不变化的设备，
              tSinceLast 会封顶在 24 天，间隔判据退化为「恒满足」——对寿命台账无实质影响，此口径未实测。
              ② 抖动计数与主计数共用 bSaturated 观测（同族计数饱和不另设码，避免凑槽，R90）。
    修订历史 :
        2026-11-16  v1.0.0  首版，R21 批次 4 入库
*)
FUNCTION_BLOCK FB_DL_SignalChangeCounter
VAR_INPUT
    bEnable         : BOOL := TRUE;      // 使能，FALSE 时冻结计数与基准，不产生新事件 / enable, FALSE freezes both the counts and the baseline
    fValue          : LREAL;             // 被监视量，如阀位 [%] / monitored value, e.g. valve position [percent]
    fDeadband       : LREAL := 1.0;      // 变化死区，同工程单位；负值按绝对值、非有限按 0 / change deadband in the same unit, negative is taken by magnitude
    tMinInterval    : TIME := T#1S;      // 最小有效变化间隔，短于此间隔的变化计入抖动 [ms] / minimum interval of an accepted change [ms]
    bReset          : BOOL;              // 上升沿清零主计数与抖动计数（不清基准）/ rising edge clears both counts but never the baseline
END_VAR
VAR_OUTPUT
    uCount          : UDINT;             // 有效变化次数，饱和后停止递增 [次] / accepted change count, stops at saturation [count]
    uChatterCount   : UDINT;             // 抖动次数（间隔不足的变化），不计入主计数 [次] / chatter count for changes inside the minimum interval [count]
    fLastAccepted   : LREAL;             // 上次被接受（或判为抖动）的值，即当前基准 [工程单位] / the baseline value, updated on every judged change [engineering unit]
    tSinceLast      : TIME;              // 距上次接受/判抖的时长，封顶 T#24D [ms] / time since the last judged change, capped at one day [ms]
    bSaturated      : BOOL;              // 任一同族计数已达上限 / at least one counter reached its upper bound
    eErr            : UDINT;             // 错误码，0=正常；16#0001_04XX 信息级 / 16#0001_03XX 故障级 / error id, 0=ok
    bError          : BOOL;              // 故障级标志 / fault flag
END_VAR
VAR
    fbElapsed       : TON;               // 间隔计时器，主体最前部无条件刷新 / interval timer, refreshed unconditionally at the top
    rtReset         : R_TRIG;            // 复位上升沿，主体最前部无条件刷新 / reset rising edge, refreshed unconditionally at the top
    bTimerKick      : BOOL;              // 计时器复位脉冲，置位后下一扫描周期 ET 归零 / reset pulse, the elapsed time restarts on the next scan
    fDeadbandEff    : LREAL;             // 生效死区，恒非负 [工程单位] / effective deadband, always non-negative [engineering unit]
    bValueFin       : BOOL;              // 当前输入是否有限 / whether the current input is finite
    bInitDone       : BOOL := FALSE;     // 首扫基准种子标志，防「0 → 当前值」的虚假首变化 / first scan seeding flag
END_VAR
VAR CONSTANT
    DL_UDINT_MAX        : UDINT := 16#FFFF_FFFF;               // 计数上限 [次] / counter upper bound [count]
    DL_TON_PT_MAX       : TIME := T#24D;                       // 计时器上限，同时是 tSinceLast 的封顶值 [ms] / timer bound and the cap of tSinceLast [ms]
    DL_LREAL_MAX_FINITE : LREAL := 1.7976931348623157E308;     // LREAL 最大有限值 [无量纲] / largest finite LREAL [dimensionless]
    DL_LREAL_ZERO       : LREAL := 0.0;                        // 零哨兵 [工程单位] / zero sentinel [engineering unit]
    DL_UDINT_ZERO       : UDINT := 0;                          // 计数零哨兵 [次] / counter zero sentinel [count]
    DL_ERR_NONE         : UDINT := 16#0000_0000;               // 无故障 / no error
END_VAR

// 段 0｜错误状态预置 / segment 0, preset the error state
eErr   := DL_ERR_NONE;                       // 预置无错误 / preset no error
bError := FALSE;                             // 预置无故障 / preset no fault

// 段 1｜定时器与边沿无条件刷新（任何 IF 之前）；踢一脚即复位 ET / segment 1, unconditional refresh, a kick restarts the elapsed time
fbElapsed( IN := NOT bTimerKick, PT := DL_TON_PT_MAX );
rtReset  ( CLK := bReset );
IF bTimerKick THEN
    bTimerKick := FALSE;                     // 复位脉冲只活一拍，本拍用完即销 / the kick lives exactly one scan
END_IF
tSinceLast := fbElapsed.ET;                  // 距上次判定变化的时长 / elapsed time since the last judged change

// 段 2｜死区参数闸：负值取绝对值、非有限按 0，不停机 / segment 2, deadband gate, never stops the machine
IF (fDeadband <> fDeadband) OR (ABS(fDeadband) > DL_LREAL_MAX_FINITE) THEN
    fDeadbandEff := DL_LREAL_ZERO;           // 非有限按零处理 / a non-finite deadband is treated as zero
    eErr   := 16#0001_039C;                  // 死区非法（故障级）/ illegal deadband, fault level
    bError := TRUE;                          // 置故障标志 / raise the fault flag
ELSIF fDeadband < DL_LREAL_ZERO THEN
    fDeadbandEff := -fDeadband;              // 负值取绝对值继续 / take the magnitude and carry on
    eErr   := 16#0001_039C;                  // 死区非法（故障级）/ illegal deadband, fault level
    bError := TRUE;                          // 置故障标志 / raise the fault flag
ELSE
    fDeadbandEff := fDeadband;               // 正常值 / a healthy value
END_IF

// 段 3｜复位沿：只清计数，不清基准 / segment 3, the reset edge clears the counts but never the baseline
IF rtReset.Q THEN
    uCount        := DL_UDINT_ZERO;          // 主计数清零 / clear the accepted count
    uChatterCount := DL_UDINT_ZERO;          // 抖动计数清零 / clear the chatter count
    bSaturated    := FALSE;                  // 解除饱和 / release the saturation flag
END_IF

// 段 4｜输入有限性判定 / segment 4, input finiteness
bValueFin := (fValue = fValue) AND (ABS(fValue) <= DL_LREAL_MAX_FINITE);   // 自比较判 NaN，幅值判 INF / self compare for NaN, magnitude for INF
IF NOT bValueFin THEN
    IF eErr = DL_ERR_NONE THEN
        eErr := 16#0001_0454;                // 输入非有限，基准保持不变（信息级）/ non-finite input, the baseline is untouched, info level
    END_IF
END_IF

// 段 5｜首扫种子：不种子就会把「0 → 当前值」记成一次虚假动作 / segment 5, first scan seeding avoids a phantom change
IF NOT bInitDone THEN
    IF bValueFin THEN
        fLastAccepted := fValue;             // 基准取首拍值 / seed the baseline with the first sample
    END_IF
    bInitDone := TRUE;                       // 种子只做一次 / seed exactly once
ELSIF bEnable AND bValueFin THEN
    // 段 6｜死区判据 + 间隔分流（核心：抖动也刷新基准）/ segment 6, deadband test and interval split, chatter updates the baseline too
    IF ABS(fValue - fLastAccepted) > fDeadbandEff THEN
        IF fbElapsed.ET >= tMinInterval THEN
            IF uCount >= DL_UDINT_MAX THEN
                bSaturated := TRUE;          // 主计数饱和 / the accepted count is saturated
                IF eErr = DL_ERR_NONE THEN
                    eErr := 16#0001_0455;    // 计数饱和（信息级）/ counter saturated, info level
                END_IF
            ELSE
                uCount := uCount + 1;        // 有效变化计数 / count the accepted change
            END_IF
        ELSE
            IF uChatterCount >= DL_UDINT_MAX THEN
                bSaturated := TRUE;          // 抖动计数饱和，同族观测 / the chatter count saturates, same observation flag
            ELSE
                uChatterCount := uChatterCount + 1;   // 间隔不足计入抖动 / a change inside the interval counts as chatter
            END_IF
        END_IF
        fLastAccepted := fValue;             // 关键：无论接受还是抖动，基准一律刷新 / the baseline is refreshed in both branches
        bTimerKick    := TRUE;               // 下一扫描周期重新起算间隔 / the interval restarts on the next scan
    END_IF
END_IF
END_FUNCTION_BLOCK

(* ---- FB_DL_SignalCrossbar8.st ---- *)
// FB_DL_SignalCrossbar8 v1.0.0
// 开源溯源：self-cleanroom / 信号路由族
(*
  道莅工业代码库 | DL_Base | FB_DL_SignalCrossbar8
  版本: 1.0.0 | 日期: 2026-11-23 | 轮次: R75
  功能: 8×8 信号交叉开关矩阵：8 路输入经路由表任意分配至 8 路输出
        （每输出独立选源 0..8，0=无源置零），同源多投允许（广播路由）
  邻件关系: 与 Mux2Ex / Mux4Ex（单选多路器）同族 —— 差异点：多路器为
            单输出 N 选 1，本件为 8 输出各 9 选 1 全交叉矩阵（含广播），
            路由自由度扩展非同义替换
  路由契约: aRoute[j] = 输出 j 的源号（0=无源/1..8=输入号），每拍执行
            刷新；越界源号按无源处理并置组态码
*)
FUNCTION_BLOCK FB_DL_SignalCrossbar8
VAR_INPUT
    aIn     : ARRAY[1..8] OF REAL;               // 8 路输入 [工程单位] / 8 inputs
    aRoute  : ARRAY[1..8] OF INT;                // 路由表（输出 j 的源号 0..8）[1] / Route table, source per output
END_VAR
VAR_OUTPUT
    aOut       : ARRAY[1..8] OF REAL;            // 8 路输出 [工程单位] / 8 outputs
    aRouteEcho : ARRAY[1..8] OF INT;             // 生效路由回显（钳位后）[1] / Effective route echo
    bValid     : BOOL;                           // 组态有效回执 [-] / Config validity receipt
    bError     : BOOL;                           // 故障标志（任一路由越界）/ Fault flag (any route out of range)
    uErrorId   : UDINT;                          // 事件码，0 = 无事件；16#0002_2201 = 路由越界 / Event code
END_VAR
VAR
    j          : INT;                            // 输出通道索引 [路] / Output channel index
    nSrc       : INT;                            // 当前源号 [1] / Current source index
END_VAR

// —— 段 0：全路径缺省 —— //
bValid := TRUE;                                  // 组态回执预置（越界路径降级）/ Validity preset
bError := FALSE;                                 // 故障预清 / Fault preset
uErrorId := 16#0000;                             // 事件码预清 / Event code preset

// —— 段 1：逐输出路由执行（源号越界按无源降级，不中断矩阵） —— //
FOR j := 1 TO 8 DO                                // 8 路输出逐一派发 / Per-output dispatch
    nSrc := aRoute[j];                            // 取该输出源号 / Source for this output
    IF (nSrc < 0) OR (nSrc > 8) THEN              // 越界源号（下标判界，R4）/ Source out of range
        aOut[j] := 0.0;                           // 无效路由输出置零（安全侧）/ Invalid route outputs zero
        aRouteEcho[j] := 0;                       // 回显钳位无源 / Echo clamped to none
        bError := TRUE;                           // 故障标志（保持型，恢复合法自动清）/ Fault flag, self-clears on valid route
        uErrorId := 16#0002_2201;                 // 信息级：路由越界 / Info level: route out of range
        bValid := FALSE;                          // 组态回执降级 / Validity degraded
    ELSIF nSrc = 0 THEN                           // 无源：输出零 / No source: zero output
        aOut[j] := 0.0;
        aRouteEcho[j] := 0;
    ELSE                                          // 合法源号 1..8：直通复制（下标判界安全）/ Valid source: pass-through
        aOut[j] := aIn[nSrc];
        aRouteEcho[j] := nSrc;
    END_IF
END_FOR
END_FUNCTION_BLOCK

(* ---- FB_DL_SignalDebounce.st ---- *)
(*==============================================================================
 * 组件名称 (Component)  : FB_DL_SignalDebounce
 * 所属子库 (Sublibrary) : DL_Base
 * 当前版本 (Version)    : 1.0.0
 * 兼容性   (Platform)   : CODESYS 3.5 / TwinCAT 3 / 汇川 InoProShop / Machine Expert
 *                         仅依赖 Standard.library（TON / R_TRIG），零厂商方言
 * 功能描述 (Function)   : 机械触点软件消抖。上升沿与下降沿确认延时独立可调，
 *                         输出消抖后稳定值 + 上升/下降单周期事件 + 消抖进行中标志。
 *                         上电首扫直接采样、不产生假边沿；延时超限自动钳位并告警；
 *                         零延时可直通；使能失效时输出直通原始值且事件清零。
 * 开源溯源 (Origin)     : 原创实现。算法思想源自 IEC 61131-3 标准定时器语义与
 *                         PLCopen Coding Guidelines 的"无条件周期刷新"约定，
 *                         未复制任何厂商私有库源码。
 * 本文件内含       : TYPE  E_DL_DebounceState（配套枚举，归属 DL_Base）
 *                    FB    FB_DL_SignalDebounce
 * 依赖     (Depends)    : 无 DL_ 内部依赖；Standard.library: TON / R_TRIG
 * 红线自检 (Redline)    : R1 ✓ 零全局变量表与外部变量引用 ｜ R2 ✓ 零物理 IO 地址直写
 *                         R3 ✓ 纯 IEC 61131-3 ｜ R4 ✓ 钳位+复位+返回值确定
 *                         R5 ✓ 全变量中英双语同行注释 ｜ R6 ✓ 五态 ENUM+CASE+ELSE
 *                         R7 ✓ 三实例主体最前部无条件刷新
 * 修订历史 (Revision)   :
 *   2026-11-14  v1.0.0  首版入库（Phase 1 冷启动 · Level 0 批次）
 *============================================================================*)

(*-----------------------------------------------------------------------------
 * 枚举: E_DL_DebounceState（归属 DL_Base，与 FB_DL_SignalDebounce 同文件）
 * 含义: 消抖状态机离散状态。数值步长留空位便于后续插态而不破坏已有工程。
 *----------------------------------------------------------------------------*)
TYPE E_DL_DebounceState :
(
    eInit     := 0,    // 上电首扫态：直接采样原始值，禁止产生任何事件 / Power-up first scan, sample directly without any event
    eStable   := 10,   // 稳定态：输出保持上一稳定值，监视输入变化 / Stable state, output holds last stable value and watches input
    eRiseWait := 20,   // 上升确认态：输入相对稳定值已变 TRUE，等待上升延时到期 / Rising confirmation, waiting for rising delay expiry
    eFallWait := 30,   // 下降确认态：输入相对稳定值已变 FALSE，等待下降延时到期 / Falling confirmation, waiting for falling delay expiry
    eFault    := 99    // 故障锁存态：非法状态或参数越界，输出回安全值，需 bReset 清除 / Latched fault, safe output, cleared by bReset
);
END_TYPE

(*==============================================================================
 * 功能块: FB_DL_SignalDebounce
 * 调用约定: 每个扫描周期无条件调用一次；bReset 上升沿重新初始化滤波器。
 * 无状态泄漏: 全部状态驻留于实例私有 VAR，零全局引用，可多实例并行。
 * 滞后披露: 输出相对输入的延迟 = 对应方向的确认延时（非固定扫描周期）。
 *============================================================================*)
FUNCTION_BLOCK FB_DL_SignalDebounce
VAR_INPUT
    bRawInput    : BOOL;              // 原始输入信号，未经消抖 / Raw input signal, not debounced
    tRiseDelay   : TIME := T#20MS;    // 上升沿确认延时 [ms]，T#0S 表示直通 / Rising confirmation delay [ms], T#0S = pass-through
    tFallDelay   : TIME := T#20MS;    // 下降沿确认延时 [ms]，T#0S 表示直通 / Falling confirmation delay [ms], T#0S = pass-through
    bEnable      : BOOL := TRUE;      // 使能标志，FALSE 时输出直通原始值 / Enable flag, FALSE bypasses output to raw input
    bReset       : BOOL;              // 复位信号，上升沿重新初始化滤波器 / Reset signal, rising edge re-initializes the filter
END_VAR
VAR_OUTPUT
    bStable      : BOOL;              // 消抖后的稳定输出 / Debounced stable output
    bRiseEvent   : BOOL;              // 稳定上升沿事件，单扫描周期脉冲 / Stable rising edge event, one-scan pulse
    bFallEvent   : BOOL;              // 稳定下降沿事件，单扫描周期脉冲 / Stable falling edge event, one-scan pulse
    bFiltering   : BOOL;              // 消抖进行中标志（输入与稳定值不一致且计时未满） / Debounce in progress flag
    bError       : BOOL;              // 故障标志，需 bReset 清除 / Fault flag, cleared by bReset
    uErrorId     : UDINT;             // 故障码，0 = 无故障 / Error code, 0 = no error
END_VAR
VAR
    fbTonRise    : TON;               // 上升确认定时器实例 / Rising confirmation timer instance
    fbTonFall    : TON;               // 下降确认定时器实例 / Falling confirmation timer instance
    fbTrigReset  : R_TRIG;            // 复位信号上升沿检测实例 / Reset rising edge detector instance
    eState       : E_DL_DebounceState; // 主状态机当前状态 / Current state of the main state machine
    bLastStable  : BOOL;              // 上一周期稳定值，仅用于边沿比较 / Previous stable value, used only for edge comparison
    tRiseClamped : TIME;              // 钳位后的上升确认延时 [ms] / Clamped rising confirmation delay [ms]
    tFallClamped : TIME;              // 钳位后的下降确认延时 [ms] / Clamped falling confirmation delay [ms]
    bNeedRise    : BOOL;              // 向上消抖请求：原始 TRUE 且稳定值 FALSE / Rise debounce request: raw TRUE while stable FALSE
    bNeedFall    : BOOL;              // 向下消抖请求：原始 FALSE 且稳定值 TRUE / Fall debounce request: raw FALSE while stable TRUE
    bRiseInstant : BOOL;              // 上升延时为零的直通快速通道标志 / Instant path flag for zero rising delay
    bFallInstant : BOOL;              // 下降延时为零的直通快速通道标志 / Instant path flag for zero falling delay
END_VAR
VAR CONSTANT
    DL_DEBOUNCE_MAX_DELAY : TIME := T#10S;  // 消抖延时上限钳位值 [s]，超限按上限执行 / Max debounce delay clamp [s], over-limit runs at clamp
END_VAR

(*------------------------------------------------------------------------------
 * 段 1｜参数钳位：延时超上限只告警不中断，保证现场不会因组态笔误停机
 *      Parameter clamping: over-limit delay only warns, never stops the machine
 *-----------------------------------------------------------------------------*)
IF tRiseDelay > DL_DEBOUNCE_MAX_DELAY THEN
    tRiseClamped := DL_DEBOUNCE_MAX_DELAY;
    bError       := TRUE;
    uErrorId     := 16#0001_0001;
ELSE
    tRiseClamped := tRiseDelay;
END_IF

IF tFallDelay > DL_DEBOUNCE_MAX_DELAY THEN
    tFallClamped := DL_DEBOUNCE_MAX_DELAY;
    bError       := TRUE;
    uErrorId     := 16#0001_0001;
ELSE
    tFallClamped := tFallDelay;
END_IF

(* 零延时判定：T#0S 必须直通，不得因 PT=0 而让输出永久不动作（边界 B4） *)
(* Zero-delay detection: T#0S must pass through, never block the output (boundary B4) *)
bRiseInstant := (tRiseClamped <= T#0S);
bFallInstant := (tFallClamped <= T#0S);

(*------------------------------------------------------------------------------
 * 段 2｜消抖需求判定：以"原始值 vs 上一周期稳定值"的偏差方向决定消抖方向
 *      Debounce request: direction derived from the deviation between raw and last stable
 *      该判定只依赖输入与上一稳定值，与状态机解耦，供下段定时器无条件使用
 *-----------------------------------------------------------------------------*)
bNeedRise := bRawInput AND NOT bStable;
bNeedFall := (NOT bRawInput) AND bStable;

(*------------------------------------------------------------------------------
 * 段 3｜无条件刷新区（红线 R7）：三个实例调用严禁进入任何 IF / CASE 分支
 *      Unconditional refresh zone (red line R7): no instance call inside IF / CASE
 *      IN 为 FALSE 时 TON 自动清零 ET，天然实现"抖动不累积计时"（边界 B8）
 *-----------------------------------------------------------------------------*)
fbTrigReset(CLK := bReset);
fbTonRise(IN := bNeedRise AND bEnable AND NOT fbTrigReset.Q, PT := tRiseClamped);
fbTonFall(IN := bNeedFall AND bEnable AND NOT fbTrigReset.Q, PT := tFallClamped);

(*------------------------------------------------------------------------------
 * 段 4｜复位处理（边界 B7）：回到 eInit 重新采样，清故障与事件
 *      Reset handling: back to eInit for re-sampling, clear fault and events
 *-----------------------------------------------------------------------------*)
IF fbTrigReset.Q THEN
    eState      := eInit;
    bError      := FALSE;
    uErrorId    := 16#0000_0000;
    bStable     := FALSE;
    bLastStable := bRawInput;
    bRiseEvent  := FALSE;
    bFallEvent  := FALSE;
    bFiltering  := FALSE;
END_IF

IF NOT bEnable THEN
    (*--------------------------------------------------------------------------
     * 段 5a｜使能失效语义（边界 B6）：直通原始值、事件清零、状态回 eInit
     *      恢复使能时由 eInit 重新采样，绝不补发禁用期间的历史边沿
     *      Disabled: bypass raw value, clear events, force eInit; no historical edge replay
     *-------------------------------------------------------------------------*)
    bStable     := bRawInput;
    bLastStable := bRawInput;
    bRiseEvent  := FALSE;
    bFallEvent  := FALSE;
    bFiltering  := FALSE;
    eState      := eInit;
ELSE
    (*--------------------------------------------------------------------------
     * 段 5b｜主状态机（红线 R6）：ENUM + CASE + ELSE 兜底
     *      Main state machine: ENUM + CASE with mandatory ELSE fallback
     *-------------------------------------------------------------------------*)
    CASE eState OF

        eInit:
            (* 首扫直接采样；bStable 与 bLastStable 同时赋值使边沿差为零（边界 B2） *)
            (* First scan samples directly; equal assignment keeps the edge difference zero *)
            bStable     := bRawInput;
            bLastStable := bRawInput;
            bRiseEvent  := FALSE;
            bFallEvent  := FALSE;
            eState      := eStable;

        eStable:
            (* 稳定监视：仅当输入偏离稳定值时才启动对应方向的确认流程 *)
            (* Stable watch: start the matching confirmation only on deviation *)
            IF bNeedRise THEN
                eState := eRiseWait;
            ELSIF bNeedFall THEN
                eState := eFallWait;
            END_IF

        eRiseWait:
            IF NOT bNeedRise THEN
                (* 输入回落：抖动被吸收，TON.IN 变 FALSE 自动清零 ET（边界 B8） *)
                (* Input bounced back: jitter absorbed, TON.IN FALSE resets ET automatically *)
                eState := eStable;
            ELSIF bRiseInstant OR fbTonRise.Q THEN
                (* 延时到期或零延时直通：确认稳定值为 TRUE *)
                (* Delay expired or zero-delay path: confirm stable value as TRUE *)
                bStable := TRUE;
                eState  := eStable;
            END_IF

        eFallWait:
            IF NOT bNeedFall THEN
                (* 输入回升：抖动被吸收，TON.IN 变 FALSE 自动清零 ET（边界 B8） *)
                (* Input recovered: jitter absorbed, TON.IN FALSE resets ET automatically *)
                eState := eStable;
            ELSIF bFallInstant OR fbTonFall.Q THEN
                (* 延时到期或零延时直通：确认稳定值为 FALSE *)
                (* Delay expired or zero-delay path: confirm stable value as FALSE *)
                bStable := FALSE;
                eState  := eStable;
            END_IF

        eFault:
            (* 故障锁存：输出回安全值 FALSE，等待 bReset 解除（边界 B9） *)
            (* Latched fault: force safe output FALSE until bReset releases it *)
            bStable := FALSE;

        ELSE
            (* 非法状态拦截：任何未定义状态一律进故障态，不做隐式恢复（边界 B9） *)
            (* Illegal state interception: any undefined state goes to fault, no implicit recovery *)
            eState   := eFault;
            bStable  := FALSE;
            bError   := TRUE;
            uErrorId := 16#0001_0005;

    END_CASE;

    (*--------------------------------------------------------------------------
     * 段 6｜边沿统一出口：只对"消抖后的稳定值"取沿（需求硬约束，边界 B5）
     *      Single edge outlet: edges are taken from the debounced stable value only
     *      放在状态机之后，任何分支改写 bStable 都只会产生一个脉冲，杜绝重发
     *-------------------------------------------------------------------------*)
    bRiseEvent := bStable AND NOT bLastStable AND NOT fbTrigReset.Q;
    bFallEvent := (NOT bStable) AND bLastStable AND NOT fbTrigReset.Q;

    (* 上一稳定值更新必须在事件计算之后，否则边沿永远为 FALSE *)
    (* Previous stable update must follow the edge evaluation, otherwise edges vanish *)
    bLastStable := bStable;

    (* 消抖进行中：处于任一确认态时为 TRUE，供 HMI 显示"滤波忙" *)
    (* Filtering busy: TRUE while in either confirmation state, for HMI display *)
    bFiltering := (eState = eRiseWait) OR (eState = eFallWait);
END_IF
END_FUNCTION_BLOCK

(* ---- FB_DL_SignalEdgeDelayEx.st ---- *)
//==============================================================================
// 功能块：FB_DL_SignalEdgeDelayEx ｜ 中文名称：边沿延迟输出（升/降沿独立延迟窗）
// 所属子库：DL_Base ｜ 版本：v1.0.0 ｜ 日期：2026-11-23
// 兼容：CODESYS V3.5+ / TwinCAT 3 / 汇川 InoProShop（纯标准库 TON）
// 功能描述：上升沿与下降沿各自独立延迟窗：bOut = (bIn AND tonRise.Q) OR
//           ((NOT bIn) AND NOT tonFall.Q)。输入置 TRUE 后经 tDelayRise 才
//           输出 TRUE；输入撤 FALSE 后经 tDelayFall 才输出 FALSE。输出待决
//           方向分别经 bPendRise / bPendFall 声明（延迟窗内 TRUE，供上层
//           做"已下令未生效"诊断）。
//           分工声明：与 FB_DL_PulseStretch（单脉冲展宽）及 TpRetrigger 族
//           互引——那两件做脉冲生成/展宽，本件只做电平沿延迟，互不替代；
//           与候选队列 FT_IMP（脉冲保持）同属脉冲定时族，本件取其"沿触发
//           电平保持"行为定义分类，不取其单脉冲语义。
// 开源溯源 (Origin)：候选队列 FT_IMP（oscatBasic，MIT 许可，
//           https://github.com/tkucic/brOscatLib/blob/main/oscatBasic/FT_IMP.st）
//           ——脉冲定时族行为定义分类参考；原名 FT_IMP → 道莅
//           FB_DL_SignalEdgeDelayEx，clean-room 独立重写（双沿独立延迟窗
//           为道莅增量，零源码行复制）
// 公开接口清单：输入 bIn / tDelayRise / tDelayFall；输出 bOut / bPendRise /
//               bPendFall / bValid
// 单位表：tDelayRise / tDelayFall [ms]，其余 BOOL 引脚无量纲
// 输入契约：bIn 为待整形原始电平；双窗参数允许为 0（对应方向直通）。
// 输出契约：bOut 为延迟后电平；bPendRise/bPendFall 为窗内瞬时待决声明
//           （每拍重算不锁存）；bValid 恒 TRUE（纯定时组合无故障级条件）。
// 错误码表：无状态机码轨（纯定时组合无故障级条件），不占用 16#0001 段码位
// 状态机：N/A（无状态机；TON ×2 每拍无条件刷新）
// 边界行为：① tDelayRise / tDelayFall 可为 0（直通，无延迟窗）；
//           ② TON 每拍无条件刷新（不入分支，红线 R7）；
//           ③ 延迟窗内撤使能无独立引脚——本件无使能门（纯信号整形件，
//             上层如需门控请在 bIn 前级串门）；
//           ④ 待决声明为窗内瞬时量，每拍重算不锁存。
// 修订历史：v1.0.0 2026-11-23 首版（R73 派单 · 批 3 · 序 14）
//==============================================================================

(*==============================================================================
 * 功能块: FB_DL_SignalEdgeDelayEx
 * 调用约定: 每个扫描周期无条件调用一次；实例状态全部驻留于 TON 实例。
 * 调用示例: edgeDelay(bIn := bRawSig, tDelayRise := T#500MS,
 *                     tDelayFall := T#200MS);
 *          bOut 替代原信号进下游判据；bPendRise/bPendFall 送上位诊断。
 * 组装说明: ① 本件无使能门，如需条件化整形请在 bIn 前级串门控合取；
 *           ② 双窗独立：tDelayRise 只作用于 TRUE 建立方向，tDelayFall
 *             只作用于 FALSE 建立方向，互不干扰；
 *           ③ 与 FB_DL_PulseStretch 分工：展宽/单脉冲用那件，电平沿
 *             延迟用本件（头注释分工声明已互引）。
 *==============================================================================*)
FUNCTION_BLOCK FB_DL_SignalEdgeDelayEx
VAR_INPUT
    bIn        : BOOL := FALSE;        // 输入信号 [—] / Input signal
    tDelayRise : TIME := T#0MS;        // 上升沿延迟窗 [ms] / Rise delay window [ms]
    tDelayFall : TIME := T#0MS;        // 下降沿延迟窗 [ms] / Fall delay window [ms]
END_VAR
VAR_OUTPUT
    bOut       : BOOL;                 // 延迟后输出 [—] / Delayed output
    bPendRise  : BOOL;                 // 上升待决声明（输入 TRUE 但窗未满）/ Rise pending, input TRUE but window open
    bPendFall  : BOOL;                 // 下降待决声明（输入 FALSE 但窗未满）/ Fall pending, input FALSE but window open
    bValid     : BOOL;                 // 输出可用标志 / Outputs usable flag
END_VAR
VAR
    tonRise    : TON;                  // 上升沿延迟定时器，每拍无条件刷新 / Rise delay timer, refreshed every scan
    tonFall    : TON;                  // 下降沿延迟定时器，每拍无条件刷新 / Fall delay timer, refreshed every scan
END_VAR

// ---- 段 1｜定时器无条件刷新（红线 R7：禁入条件分支）----
tonRise(IN := bIn,  PT := tDelayRise); // 上升窗计时随输入断续 / Rise timer input follows the signal
tonFall(IN := NOT bIn, PT := tDelayFall); // 下降窗计时随输入反相断续 / Fall timer input follows the inverted signal

// ---- 段 2｜输出主体：双沿门控合成（升沿等 tonRise.Q，降沿借 tonFall 未满）----
bOut := (bIn AND tonRise.Q) OR ((NOT bIn) AND (NOT tonFall.Q)); // 双沿独立延迟合成 / Dual-edge independent delay blend

// ---- 段 3｜待决声明：窗内瞬时量每拍重算（诊断用，不锁存）----
bPendRise := bIn AND (NOT tonRise.Q); // 上升窗未满待决 / Rise pending while window open
bPendFall := (NOT bIn) AND (NOT tonFall.Q); // 下降窗未满待决 / Fall pending while window open
bValid := TRUE;                       // 纯定时组合恒可用 / Pure timing combinational, always usable
END_FUNCTION_BLOCK

(* ---- FB_DL_SignalFreeze.st ---- *)
(*==============================================================================
 * 组件名称 (Component)  : FB_DL_SignalFreeze
 * 所属子库 (Sublibrary) : DL_Base
 * 当前版本 (Version)    : 1.0.0
 * 兼容性   (Platform)   : CODESYS 3.5 / TwinCAT 3 / 汇川 InoProShop / Machine Expert
 *                         仅依赖 Standard.library（TON / R_TRIG），零厂商方言
 * 来源标签 (Source)     : self-std（防御性新增线）
 * 功能描述 (Function)   : 坏值冻结保持：连续量输入出现 NaN / Inf / 越合理性域时，
 *                         输出保持上一次有效值（绝不把坏值搬到下游），并累计冻结
 *                         时长；冻结时长超过 tFreezeMax 即判「信号源已死」锁存告警。
 *                         有效输入回来时：输出无扰切回实时值，冻结计时清零。
 * 分工互引 (Boundary)   : ① FB_DL_SignalHoldResume —— 由**外部命令 bHold** 决定
 *                         保持还是恢复（人工/工艺保持），不判信号真伪；
 *                         ② FB_DL_SignalFrozenDetect —— 判「信号数值长期不变」的
 *                         冻结故障（上游诊断）；③ 本件由**坏值**驱动自动保持 +
 *                         冻结时长告警，三件语义互不重叠，禁互相替代。
 * 边界与语义披露 (Boundary disclosure) :
 *   1) 合理性域 [fLowLim, fHighLim] 为闭区间；fLowLim > fHighLim 属组态非法，
 *      锁存至复位沿 + 组态改对（R152 解除路径自证）。
 *   2) 坏值判定三判据全枚举（R272）：NaN 自反 `x <> x`、Inf 差自减
 *      `(x − x) <> (x − x)`、幅值兜底 `ABS(x) >= 1.0E30`。禁用单一近似阈值。
 *   3) 坏值期输出恒为**上一次有效值**（fHold 只在有效样本上刷新），因此输出永远
 *      有限；下游无需再做非有限防护（但本件仍不承诺输出在域内——保持值属于
 *      历史有效值，域闸变更后可能落在新域外，这是刻意保留的证据语义）。
 *   4) 冻结时长超限为**故障级锁存**：解除 = 复位沿 AND 本拍输入有效（信号已恢复），
 *      未恢复时复位沿不作解除（防复位即掩盖断线）。
 *   5) 冻结告警不是动作输出：本件只上报，不切断工艺（切断归使用侧联锁件）。
 * 故障码表 (Error codes) :
 *   16#0001_03FC [故障级] 组态非法（合理性域反向 / 冻结上限 <= T#0S），不冻结不告警
 *                 反证：禁用与组态非法都表现为「输出恒等输入」，现有输出不可区分。
 *   16#0001_03FD [故障级] 冻结时长超限（信号源疑似失效），锁存至复位沿 + 输入恢复
 *                 反证：持续坏值与「信号源恰好长时间恒定为某有效值」输出组合相同，
 *                 无码则该故障对 HMI 完全不可见。
 *   16#0001_04FD [信息级] 本拍进入坏值冻结保持（bFrozen 同源可查）
 *                 反证：冻结与「输入稳定不变」输出组合相同；单拍级事件事实需入流水。
 * 码位总账 (Code ledger) : 16#0001_03FC / 03FD 用 ｜ 16#0001_04FD 用
 * 依赖     (Depends)    : 无 DL_ 内部依赖；Standard.library: TON / R_TRIG
 * 红线自检 (Redline)    : R1 ✓ 零全局变量与 VAR_EXTERNAL ｜ R2 ✓ 零 %I/%Q 物理地址
 *                         R3 ✓ 纯 IEC 61131-3 ｜ R4 ✓ 非有限三判 / 无除法 / 域闸全枚举
 *                         R5 ✓ 全变量中英双语同行注释 ｜ R6 ✓ 四态 ENUM + CASE + ELSE
 *                         R7 ✓ 一沿一计时主体最前部无条件刷新
 * 修订历史 (Revision)   :
 *   2026-11-22  v1.0.0  首版入库（R69 构建轮 · 批 2 · N7）
 *============================================================================*)

(*-----------------------------------------------------------------------------
 * 枚举: E_DL_FreezeState（归属 DL_Base，与 FB_DL_SignalFreeze 同文件）
 *----------------------------------------------------------------------------*)
TYPE E_DL_FreezeState :
(
    eIdle   := 0,     // 未使能：输出恒等于输入（不保持）/ Disabled, output mirrors the input
    ePass   := 10,    // 实时直通：输入有效 / Live pass-through, input valid
    eFrozen := 20,    // 坏值冻结：输出保持上次有效值 / Frozen, outputs the last valid value
    eAlarm  := 99     // 冻结超限锁存：输出仍保持，需人工复位 / Frozen too long, latched
);
END_TYPE

(*==============================================================================
 * 功能块: FB_DL_SignalFreeze
 * 调用约定: 每个扫描周期无条件调用一次；bReset 为上升沿语义。
 *============================================================================*)
FUNCTION_BLOCK FB_DL_SignalFreeze
VAR_INPUT
    fIn         : REAL;                  // 连续量输入 [工程单位] / continuous input [engineering unit]
    fLowLim     : REAL := -1.0E6;        // 合理性域下限（含）[工程单位] / plausibility floor, inclusive
    fHighLim    : REAL := 1.0E6;         // 合理性域上限（含）[工程单位] / plausibility ceiling, inclusive
    tFreezeMax  : TIME := T#5S;          // 冻结时长告警上限 [s]，<= T#0S 组态非法 / freeze duration ceiling [s]
    bEnable     : BOOL := TRUE;          // 使能；FALSE 时输出恒等输入（降级已声明）/ enable, FALSE mirrors the input
    bReset      : BOOL;                  // 上升沿：清冻结超限锁存（须输入已恢复）/ rising edge clears the freeze latch
END_VAR
VAR_OUTPUT
    fOut        : REAL;                  // 输出（坏值期 = 上次有效值）[工程单位] / output, last valid while frozen
    bFrozen     : BOOL;                  // 本拍处于坏值冻结保持 / frozen this scan
    tFrozenDur  : TIME;                  // 当前冻结已持续时长 [s] / current freeze duration [s]
    bFreezeAlarm: BOOL;                  // 冻结时长超限锁存（人工复位解除）/ freeze duration exceeded, latched
    bInputValid : BOOL;                  // 本拍输入有效（域内且有限）/ input valid this scan
    bError      : BOOL;                  // 故障标志（组态 / 冻结超限锁存）/ fault flag
    uErrorId    : UDINT;                 // 故障码，0 = 无故障 / error code, 0 = none
    eState      : E_DL_FreezeState;      // 当前状态（供 HMI 诊断）/ current state for HMI diagnosis
END_VAR
VAR
    fbTrigReset : R_TRIG;                // 复位沿检测实例 / reset edge detector
    tonFreeze   : TON;                   // 冻结时长计时实例 / freeze duration timer
    eStateInt   : E_DL_FreezeState;      // 主状态机内部当前态 / internal state machine state
    fHold       : REAL;                  // 上次有效值保持槽 [工程单位] / hold slot of the last valid value
    bInValidT   : BOOL;                  // 本拍输入有效（含域闸）/ input valid this scan including the domain gate
    bCfgBad     : BOOL;                  // 本拍组态非法 / config illegal this scan
    bCfgLatch   : BOOL;                  // 组态锁存（复位沿 + 组态改对解除）/ config latch
    bAlarmInt   : BOOL;                  // 冻结超限锁存内部副本 / internal freeze alarm latch
    bErrorInt   : BOOL;                  // 本拍故障置位累加（出口归并）/ fault set accumulator of this scan
    bFirstScan  : BOOL := TRUE;          // 上电首扫标志 / first-scan flag
END_VAR
VAR CONSTANT
    DL_SF_FIN_LIM : REAL := 1.0E30;      // REAL 幅值兜底判界 / REAL magnitude bound as the last line
    DL_SF_NO_ALARM : REAL := 0.0;        // 有限零点常量（首扫落零）[工程单位] / finite zero constant for first scan
END_VAR

(*------------------------------------------------------------------------------
 * 段 1｜无条件刷新区（红线 R7）：一沿一计时位于主体最前部
 *      Unconditional refresh: one edge and one timer at the very top
 *-----------------------------------------------------------------------------*)
fbTrigReset(CLK := bReset);
tonFreeze(IN := (eStateInt = E_DL_FreezeState.eFrozen), PT := tFreezeMax);

(*------------------------------------------------------------------------------
 * 段 2｜上电首扫：保持槽落有限零点（禁用未初始化量参与下游）/ first-scan init
 *-----------------------------------------------------------------------------*)
IF bFirstScan THEN
    eStateInt  := E_DL_FreezeState.eIdle;
    fHold      := DL_SF_NO_ALARM;
    bAlarmInt  := FALSE;
    bFirstScan := FALSE;
END_IF

(* 段 3｜每拍预清（FB32-1）：单拍标志，禁入锁存 / per-scan preset, single-scan flags only *)
bErrorInt := FALSE;

(*------------------------------------------------------------------------------
 * 段 4｜组态域闸（R151）：合理性域反向 / 冻结上限非正即非法，锁存至复位沿
 *      Config gate: reversed plausibility interval or non-positive ceiling
 *      解除路径（R152 自证）：复位沿 AND 组态已改对
 *-----------------------------------------------------------------------------*)
bCfgBad := (fLowLim > fHighLim) OR (fLowLim <> fLowLim) OR (fHighLim <> fHighLim)
           OR (tFreezeMax <= T#0S);

IF bCfgBad THEN
    bCfgLatch := TRUE;
END_IF
IF fbTrigReset.Q AND (NOT bCfgBad) THEN
    bCfgLatch := FALSE;              // 组态锁存解除 / config latch cleared
    uErrorId  := 16#0000_0000;       // 码位随解除归零 / code cleared with the latch
END_IF
IF bCfgLatch THEN
    uErrorId  := 16#0001_03FC;       // 故障级：组态非法 / fault: illegal configuration
    bErrorInt := TRUE;               // R45 配对 / paired with the code
END_IF

(*------------------------------------------------------------------------------
 * 段 5｜坏值三判（R272）：NaN 自反 / Inf 差自减 / 幅值兜底，再并合理性域
 *      Bad-value triage: NaN, Inf and the plausibility interval
 *-----------------------------------------------------------------------------*)
bInValidT := (NOT (fIn <> fIn))
             AND (NOT ((fIn - fIn) <> (fIn - fIn)))
             AND (ABS(fIn) < DL_SF_FIN_LIM)
             AND (fIn >= fLowLim) AND (fIn <= fHighLim)
             AND bEnable
             AND (NOT bCfgLatch);

(*------------------------------------------------------------------------------
 * 段 6｜主状态机（红线 R6）：ENUM + CASE + ELSE 兜底
 *      拍 N 进入：本拍坏值 -> eFrozen 并保持 fHold；本拍行为：不刷新 fHold；
 *      拍 N+1 转出：输入恢复有效即回 ePass 并清冻结计时（无扰切回实时值）
 *-----------------------------------------------------------------------------*)
CASE eStateInt OF

    E_DL_FreezeState.eIdle:
        IF bEnable AND (NOT bCfgLatch) THEN
            eStateInt := E_DL_FreezeState.ePass;    // 使能且组态合法才进入直通 / enabled and configured
        END_IF

    E_DL_FreezeState.ePass:
        IF (NOT bEnable) OR bCfgLatch THEN
            eStateInt := E_DL_FreezeState.eIdle;    // 失能 / 组态非法即退出 / disable or config fault
        ELSIF NOT bInValidT THEN
            eStateInt := E_DL_FreezeState.eFrozen;  // 坏值：进冻结保持 / bad value, start holding
            uErrorId  := 16#0001_04FD;              // 信息级：进入冻结保持 / info: frozen hold entered
        END_IF

    E_DL_FreezeState.eFrozen:
        IF (NOT bEnable) OR bCfgLatch THEN
            eStateInt := E_DL_FreezeState.eIdle;
        ELSIF bInValidT THEN
            eStateInt := E_DL_FreezeState.ePass;    // 输入恢复：无扰切回实时 / recovered, back to live
        ELSIF bAlarmInt THEN
            eStateInt := E_DL_FreezeState.eAlarm;   // 冻结超限：迁告警态驻留 / frozen too long
        END_IF

    E_DL_FreezeState.eAlarm:
        (* 输出仍保持上次有效值（不因告警改口径）；解除 = 复位沿 AND 输入已恢复 *)
        IF fbTrigReset.Q AND bInValidT AND (NOT bCfgBad) THEN
            bAlarmInt  := FALSE;                    // 冻结超限锁存解除 / alarm latch cleared
            uErrorId   := 16#0000_0000;
            eStateInt  := E_DL_FreezeState.ePass;   // 直接回直通（本拍输入已有效）/ straight back to pass-through
        ELSIF (NOT bEnable) OR bCfgLatch THEN
            eStateInt  := E_DL_FreezeState.eIdle;
        END_IF

    ELSE
        (* 非法状态拦截：迁兜底态并锁存上报 / illegal state interception *)
        eStateInt := E_DL_FreezeState.eAlarm;
        bAlarmInt := TRUE;
        uErrorId  := 16#0001_03FD;
        bErrorInt := TRUE;

END_CASE;

(*------------------------------------------------------------------------------
 * 段 7｜保持槽刷新与冻结计时消化（保持槽只在有效样本上写）
 *      Hold slot refresh and freeze timer digestion
 *-----------------------------------------------------------------------------*)
IF bInValidT THEN
    fHold := fIn;                    // 有效样本刷新保持槽 [工程单位] / refresh the hold slot
END_IF

IF tonFreeze.Q AND (NOT bAlarmInt) THEN
    bAlarmInt := TRUE;               // 冻结超限锁存 / freeze alarm latched
    uErrorId  := 16#0001_03FD;       // 故障级：冻结时长超限 / fault: freeze duration exceeded
    bErrorInt := TRUE;               // R45 配对 / paired with the code
    eStateInt := E_DL_FreezeState.eAlarm;
END_IF

(*------------------------------------------------------------------------------
 * 段 8｜输出单一出口（范式 P-05）：输出恒为保持槽（有限），坏值永不外泄
 *      Single output exit: the output is always the finite hold slot
 *-----------------------------------------------------------------------------*)
fOut        := fHold;                                      // 输出 = 上次有效值 [工程单位] / output equals the last valid value
bFrozen     := (eStateInt = E_DL_FreezeState.eFrozen) OR (eStateInt = E_DL_FreezeState.eAlarm);
tFrozenDur  := tonFreeze.ET;                               // 当前冻结时长 [s] / current freeze duration
bFreezeAlarm := bAlarmInt;                                 // 超限锁存直出 / alarm latch straight out
bInputValid := bInValidT;                                  // 本拍有效性直出 / validity straight out
bError      := bErrorInt OR (eStateInt = E_DL_FreezeState.eAlarm) OR bCfgLatch;
eState      := eStateInt;
END_FUNCTION_BLOCK

(* ---- FB_DL_SignalFrozenDetect.st ---- *)
(*
    组件名称 : FB_DL_SignalFrozenDetect
    所属子库 : DL_Base
    当前版本 : 1.0.0
    兼 容 性 : CODESYS V3.5+ / TwinCAT 3 / 汇川 InoProShop；仅依赖 Standard.library
    功能描述 : 信号冻结检测，窗内极差小于死区即判传感器卡死；NE107 的 eCheckFunction（功能自检）判据原子。
              取舍 ①：窗内只跟踪极值（fMin / fMax 增量更新），不开数组 —— 观察窗可能长达数分钟，
              按扫描周期存样本要几千个 LREAL，用极差判冻结只需两个数，内存与扫描开销都降到常数。
              取舍 ②：非有限输入不推进窗、不更新极值 —— NaN / INF 不是「冻结」也不是「变化」，
              把它们塞进极值会让整窗作废；本件暂停窗并发信息码，同时用第二只定时器累计「连续非有限」时长，
              超窗即判信号失效（03A3），与「冻结」严格区分：一个是传感器卡住，一个是信号链断了。
              取舍 ③：暂停窗的实现是定时器失电复位（保守侧）—— 严格「暂停」需要保存已累计时长，
              那就要引入额外时基量并面对漂移；宁可让窗重新起算，也只在「推迟判定」这个安全方向上让步。
              取舍 ④：解冻条件用「本拍增量超死区」而不是「极差超死区」—— 极差在窗满之后已经没用了，
              只有新增变化才说明传感器又开始动了，判据必须落在增量上。
    开源溯源 : T2-8 NE107 语义（eCheckFunction 需要功能自检判据）+ T0-1 变体线。判据、阈值、码位、；本件为道莅 clean-room 防御性实现（仅借 NE107 eCheckFunction 判据语义，零代码复制）。
              状态组织 100% 自有，零代码行与注释复制。
    本文件内含 : FUNCTION_BLOCK FB_DL_SignalFrozenDetect（单 POU，无配套类型）
    依 赖 : 无 DL_ 内部依赖；Standard.library: TON / R_TRIG
    红线自检 : R1 ✓ 零全局变量与外部变量 ｜ R2 ✓ 零物理 IO 地址
              R3 ✓ 纯 IEC 61131-3 ｜ R4 ✓ 参数闸 + 非有限闸 + 窗定时器 + 失效时长闸 + 极差容差判据
              R5 ✓ 全变量中英双语同行注释 ｜ R6 N/A 无顺序状态机（判据累加型），头注释已写明理由
              R7 ✓ 三只 TON 与 R_TRIG 全部在主体最前部无条件刷新，位于任何 IF 之外
              R8 ✓ 窗口缺省值、容差、计时上限全常量化
    错误码   : 16#0001_0458 [信息级] 输入非有限，窗暂停且极值不更新，bError = FALSE
               16#0001_0459 [信息级] 窗内极差为零（完全无抖动），bError = FALSE
               16#0001_03A2 [故障级] 窗口时长或死区非法，已钳缺省值继续，bError = TRUE
               16#0001_03A3 [故障级] 连续非有限超过一个窗口，判信号失效（区别于冻结），bError = TRUE
               16#0001_03A4 [故障级] 预留禁用（不得挪用）
    码位总账 : 16#0001_0458 用 / 16#0001_0459 用 ｜ 16#0001_03A2 用 / 16#0001_03A3 用 / 16#0001_03A4 预留
    遗留假设 : ① tFrozenFor 由一只 TON 的 ET 提供，封顶 T#24H；冻结超过 24 小时的极端工况下该值封顶，
              判定本身不受影响（bFrozen 已锁存）。此口径未实测。
              ② 窗定时器在非有限拍失电复位（保守侧），已在取舍 ③ 声明；若工艺要求「严格暂停」，
              应改由调用方注入 tDelta 自建计时，属后续变体，不在本版范围。
    修订历史 :
        2026-11-16  v1.0.0  首版，R21 批次 4 入库
*)
FUNCTION_BLOCK FB_DL_SignalFrozenDetect
VAR_INPUT
    bEnable         : BOOL := TRUE;      // 使能，FALSE 时窗停走但不改变已锁存的冻结判定 / enable, FALSE stops the window but keeps the latched verdict
    fValue          : LREAL;             // 被监视量，同死区工程单位 [工程单位] / monitored value in the deadband unit [engineering unit]
    fMoveEps        : LREAL := 0.05;     // 判定「有变化」的最小增量，负值钳缺省 [工程单位] / smallest increment that counts as movement [engineering unit]
    tWindow         : TIME := T#30S;     // 观察窗时长，≤ 0 时钳缺省 [ms] / observation window length, clamped when not positive [ms]
    bReset          : BOOL;              // 上升沿清冻结判定与窗 / rising edge clears the verdict and the window
END_VAR
VAR_OUTPUT
    bFrozen         : BOOL;              // 冻结判定，锁存至输入恢复变化或复位 / frozen verdict latched until movement or reset
    tFrozenFor      : TIME;              // 已冻结时长，封顶 T#24H [ms] / time already frozen, capped at one day [ms]
    fSpan           : LREAL;             // 窗内极差 = 最大 − 最小 [工程单位] / span inside the window [engineering unit]
    bInvalidInput   : BOOL;              // 输入非有限标志（与冻结区分）/ non-finite input flag, distinct from the frozen verdict
    eErr            : UDINT;             // 错误码，0=正常；16#0001_04XX 信息级 / 16#0001_03XX 故障级 / error id, 0=ok
    bError          : BOOL;              // 故障级标志 / fault flag
END_VAR
VAR
    fbWindow        : TON;               // 观察窗定时器，主体最前部无条件刷新 / window timer, refreshed unconditionally at the top
    fbInvalid       : TON;               // 连续非有限时长定时器，主体最前部无条件刷新 / invalid duration timer, refreshed unconditionally at the top
    fbFrozen        : TON;               // 冻结时长定时器，主体最前部无条件刷新 / frozen duration timer, refreshed unconditionally at the top
    rtReset         : R_TRIG;            // 复位上升沿，主体最前部无条件刷新 / reset rising edge, refreshed unconditionally at the top
    bWinKick        : BOOL;              // 窗复位脉冲，置位后下一扫描周期窗重新起算 / window restart pulse, effective on the next scan
    fMinVal         : LREAL;             // 窗内最小值 [工程单位] / minimum inside the window [engineering unit]
    fMaxVal         : LREAL;             // 窗内最大值 [工程单位] / maximum inside the window [engineering unit]
    fPrevValue      : LREAL;             // 上一拍输入，用于增量判据 [工程单位] / previous sample used by the movement test [engineering unit]
    fMoveEpsEff     : LREAL;             // 生效死区，恒非负 [工程单位] / effective deadband, always non-negative [engineering unit]
    tWindowEff      : TIME;              // 生效窗口时长 [ms] / effective window length [ms]
    bValueFin       : BOOL;              // 当前输入是否有限 / whether the current input is finite
    bMoved          : BOOL;              // 本拍是否检出真实变化 / whether real movement was detected this scan
    bInitDone       : BOOL := FALSE;     // 首扫极值种子标志 / first scan seeding flag
END_VAR
VAR CONSTANT
    DL_MOVE_EPS_DEF     : LREAL := 0.05;                       // 死区缺省值 [工程单位] / default deadband [engineering unit]
    DL_WINDOW_DEF       : TIME := T#30S;                       // 窗口缺省值 [ms] / default window length [ms]
    DL_TIME_ZERO        : TIME := T#0S;                        // 零时长哨兵 [ms] / zero duration sentinel [ms]
    DL_FROZEN_PT_MAX    : TIME := T#24H;                       // 冻结时长上限 [ms] / frozen duration bound [ms]
    DL_LREAL_MAX_FINITE : LREAL := 1.7976931348623157E308;      // LREAL 最大有限值 [无量纲] / largest finite LREAL [dimensionless]
    DL_LREAL_ZERO       : LREAL := 0.0;                        // 零哨兵 [工程单位] / zero sentinel [engineering unit]
    DL_FLOAT_EPS        : LREAL := 1.0E-12;                    // 极差判零容差，禁用 = 判等 [工程单位] / tolerance of the zero span test [engineering unit]
    DL_ERR_NONE         : UDINT := 16#0000_0000;               // 无故障 / no error
END_VAR

// 段 0｜错误状态预置 / segment 0, preset the error state
eErr   := DL_ERR_NONE;                    // 预置无错误 / preset no error
bError := FALSE;                          // 预置无故障 / preset no fault
bMoved := FALSE;                          // 本拍未检出变化 / no movement detected this scan

// 段 1｜参数闸：窗口与死区非法时钳缺省值继续 / segment 1, parameter gate with clamping
IF tWindow <= DL_TIME_ZERO THEN
    tWindowEff := DL_WINDOW_DEF;          // 钳缺省窗口 / clamp to the default window
    eErr   := 16#0001_03A2;               // 参数非法（故障级）/ illegal parameter, fault level
    bError := TRUE;                       // 置故障标志 / raise the fault flag
ELSE
    tWindowEff := tWindow;                // 正常值 / a healthy value
END_IF
IF (fMoveEps <> fMoveEps) OR (ABS(fMoveEps) > DL_LREAL_MAX_FINITE) OR (fMoveEps < DL_LREAL_ZERO) THEN
    fMoveEpsEff := DL_MOVE_EPS_DEF;       // 非有限或负值钳缺省 / a non-finite or negative deadband falls back to the default
    eErr   := 16#0001_03A2;               // 参数非法（故障级）/ illegal parameter, fault level
    bError := TRUE;                       // 置故障标志 / raise the fault flag
ELSE
    fMoveEpsEff := fMoveEps;              // 正常值 / a healthy value
END_IF

// 段 2｜三只定时器与边沿无条件刷新（任何 IF 之前）/ segment 2, three timers and the edge refreshed unconditionally
bValueFin := (fValue = fValue) AND (ABS(fValue) <= DL_LREAL_MAX_FINITE);   // 有限性判定 / finiteness test
bInvalidInput := NOT bValueFin;                                            // 对外暴露非有限标志 / publish the non-finite flag
fbWindow ( IN := bEnable AND bValueFin AND NOT bWinKick, PT := tWindowEff );
fbInvalid( IN := bInvalidInput,                          PT := tWindowEff );
fbFrozen ( IN := bFrozen AND bEnable,                    PT := DL_FROZEN_PT_MAX );
rtReset  ( CLK := bReset );
IF bWinKick THEN
    bWinKick := FALSE;                    // 复位脉冲只活一拍，本拍用完即销 / the restart pulse lives exactly one scan
END_IF
tFrozenFor := fbFrozen.ET;                // 已冻结时长 / elapsed frozen time

// 段 3｜非有限处理：不更新极值、不推进窗，并累计失效时长 / segment 3, non-finite handling, the window is not advanced
IF bInvalidInput THEN
    IF eErr = DL_ERR_NONE THEN
        eErr := 16#0001_0458;             // 输入非有限，窗暂停（信息级）/ non-finite input, the window pauses, info level
    END_IF
    IF fbInvalid.Q THEN
        eErr   := 16#0001_03A3;           // 连续非有限超一个窗口，判信号失效（故障级）/ invalid for a full window, fault level
        bError := TRUE;                   // 置故障标志 / raise the fault flag
    END_IF
END_IF

// 段 4｜首扫种子：极值与上拍值同时落定，防「0 → 当前值」被当成一次变化 / segment 4, first scan seeding
IF NOT bInitDone THEN
    IF bValueFin THEN
        fMinVal    := fValue;             // 最小值种子 / seed the minimum
        fMaxVal    := fValue;             // 最大值种子 / seed the maximum
        fPrevValue := fValue;             // 上拍值种子 / seed the previous sample
    END_IF
    bInitDone := TRUE;                    // 种子只做一次 / seed exactly once
    fSpan     := DL_LREAL_ZERO;           // 首扫极差为 0 / the span starts at zero
ELSIF bValueFin THEN
    // 段 5｜极值增量更新 / segment 5, incremental extreme tracking
    IF fValue < fMinVal THEN
        fMinVal := fValue;                // 刷新最小 / refresh the minimum
    END_IF
    IF fValue > fMaxVal THEN
        fMaxVal := fValue;                // 刷新最大 / refresh the maximum
    END_IF
    fSpan := fMaxVal - fMinVal;           // 窗内极差 / the span inside the window

    // 段 6｜增量判据：本拍真实变化即解冻、清窗、重种极值 / segment 6, movement releases the verdict and restarts the window
    IF ABS(fValue - fPrevValue) > fMoveEpsEff THEN
        bMoved := TRUE;                   // 检出真实变化 / real movement detected
    END_IF
    fPrevValue := fValue;                 // 上拍值无条件刷新 / the previous sample is always refreshed
    IF bMoved THEN
        bFrozen := FALSE;                 // 解冻 / release the verdict
        bWinKick := TRUE;                 // 窗从下一扫描周期重新起算 / the window restarts on the next scan
        fMinVal := fValue;                // 极值以当前值重种 / re-seed the extremes with the current sample
        fMaxVal := fValue;                // 极值基准取当前值 / extrema baseline takes current value
        fSpan   := DL_LREAL_ZERO;         // 极差归零 / reset the span
    ELSE
        // 段 7｜冻结判定：窗满且极差小于死区 / segment 7, frozen verdict when the window is full and the span is tiny
        IF fbWindow.Q AND (fSpan < fMoveEpsEff) THEN
            bFrozen := TRUE;              // 锁存冻结判定 / latch the frozen verdict
        END_IF
        IF (ABS(fSpan) < DL_FLOAT_EPS) AND (eErr = DL_ERR_NONE) THEN
            eErr := 16#0001_0459;         // 窗内极差为零（信息级）/ zero span inside the window, info level
        END_IF
    END_IF
END_IF

// 段 8｜复位沿：清判定与窗（放在判定之后，保证本拍先诊断再清）/ segment 8, reset edge after the diagnosis
IF rtReset.Q THEN
    bFrozen := FALSE;                     // 清冻结判定 / clear the verdict
    bWinKick := TRUE;                     // 窗重新起算 / restart the window
    fSpan := DL_LREAL_ZERO;               // 极差归零 / reset the span
    IF bValueFin THEN
        fMinVal := fValue;                // 极值重种 / re-seed the extremes
        fMaxVal := fValue;                // 极值基准取当前值 / extrema baseline takes current value
    END_IF
END_IF
END_FUNCTION_BLOCK

(* ---- FB_DL_SignalHoldResume.st ---- *)
(*==============================================================================
 * 组件名称 (Component)  : FB_DL_SignalHoldResume
 * 所属子库 (Sublibrary) : DL_Base
 * 当前版本 (Version)    : 1.0.0
 * 兼容性   (Platform)   : CODESYS 3.5+ / TwinCAT 3 / 汇川 InoProShop / 施耐德 Machine Expert
 *                         仅依赖 Standard.library（R_TRIG / F_TRIG），零厂商私有库
 * 功能描述 (Function)   : 8 路信号快照锁存/恢复：bHold 上升沿将 8 路实时输入
 *                         abSignal[0..7] 拍照锁存到锁存副本 abSnap；bHold=TRUE
 *                         期间输出 abOut 保持锁存副本（实时变化不穿透）；bHold
 *                         下降沿（恢复沿）输出无扰切回实时值，并逐通道做
 *                         「锁存副本 vs 实时值」一致性校验：不一致通道记入
 *                         uChgMask 位图与信息码 eResumeDiff（信息级，不置 bError）。
 * 接口     (Interface)  : 输入 abSignal 8 路实时信号数组、bHold 保持/恢复命令；
 *                         输出 abOut 8 路输出（保持期=锁存副本，恢复期=实时值）、
 *                         abSnap 锁存副本透读（诊断用）、uChgMask 恢复沿不一致
 *                         位图（bit i 对应通道 i，恢复沿单拍更新）、bHolding
 *                         保持中指示、eErrCode 信息码、bError 故障标志
 *                         （本件无故障级条件，恒 FALSE，出口保留契约位）。
 * 边界     (Boundary)   : ① **属主边界（写死）：本件只做快照锁存与恢复校验，
 *                         不判定信号真伪、不接管联锁**；信号质量诊断归
 *                         `FB_DL_SignalQualify`。
 *                         ② 锁存判定只读锁存副本（abSnap），禁止读实时数组替代
 *                         （锁存副本与实时镜像不得混用，派单红线）。
 *                         ③ 恢复沿校验用锁存副本与当拍实时值比较；uChgMask 在
 *                         非恢复沿拍保持上拍值（诊断锁存语义，非单拍抹除）。
 *                         ④ 两沿实例（R_TRIG/F_TRIG）段 0 无条件周期调用（R6）。
 *                         ⑤ 通道数定长 8（常量），无数组越界路径。
 *                         ⑥ 零全局耦合（无 GVL / VAR_EXTERNAL / 物理地址）。
 * 分工声明 (Scope)      : 与 `FB_DL_SignalFrozenDetect` 分工：信号冻结检测归那件、
 *                         快照锁存/恢复归本件；与 `FB_DL_BitShiftRegister` 分工：
 *                         移位 ≠ 快照。
 * 来源标签 (Source Tag) : 自研线（快照锁存语义为道莅防御性实现）
 * 码表     (Codes)      : 本件不占用任何全局数字码位。出口为 BOOL 数组 + WORD
 *                         位图 + ENUM 信息码；数字码位待主控收口阶段统一派号。
 * 红线自检 (Redline)    : R1 ✓ 零 GVL/VAR_EXTERNAL ｜ R2 ✓ 零 %I/%Q/%M ｜ R3 ✓ 纯 IEC 61131-3
 *                         R4 ✓ 锁存副本/实时镜像分用 ｜ R5 ✓ 声明逐行同行双语注释
 *                         R6 N/A（无 ENUM 状态机） ｜ R7 ✓ 一 R_TRIG 一 F_TRIG 段 0 无条件刷新
 * 修订历史 (Revision)   : 2026-11-20  v1.0.0  R50 首版（批次 1 · 序号 2）
 * 验收向量 (Acceptance) : ① 实时 [F,T,F,F,F,F,F,F] 时 bHold 上升沿 → abSnap=
 *                         [F,T,...]，随后 abSignal[1] 变 F：保持期 abOut 仍
 *                         [F,T,...]（变化不穿透），bHolding=TRUE；
 *                         ② bHold 下降沿：abOut 切回实时 [F,F,...]，通道 1
 *                         锁存副本 T ≠ 实时 F → uChgMask.bit1=1，
 *                         eErrCode=eResumeDiff（信息级）；
 *                         ③ 锁存副本与实时全一致时恢复 → uChgMask=0，
 *                         eErrCode=eOk。
 *==============================================================================*)

(*-----------------------------------------------------------------------------
 * 枚举: E_DL_ShrErr（信息码；本件无故障级条件，信息级不置 bError）
 *----------------------------------------------------------------------------*)
TYPE E_DL_ShrErr :
(
    eOk         := 0,   // 恢复沿锁存副本与实时一致 / Snapshot matches live at resume
    eResumeDiff := 1    // 信息级：恢复沿存在不一致通道（见 uChgMask） / Info: mismatch channels at resume, see uChgMask
);
END_TYPE

FUNCTION_BLOCK FB_DL_SignalHoldResume
VAR_INPUT
    abSignal : ARRAY[0..7] OF BOOL;   // 8 路实时输入信号 [-] / Eight live input signals
    bHold    : BOOL := FALSE;         // 保持/恢复命令（上升沿拍照，下降沿恢复） [-] / Hold command, rising edge snapshots
END_VAR
VAR_OUTPUT
    abOut    : ARRAY[0..7] OF BOOL;   // 8 路输出（保持期=锁存副本，恢复期=实时） [-] / Eight outputs
    abSnap   : ARRAY[0..7] OF BOOL;   // 锁存副本透读（诊断用） [-] / Latched snapshot for diagnostics
    uChgMask : WORD;                  // 恢复沿不一致位图（bit i=通道 i） [-] / Mismatch bitmap at resume edge
    bHolding : BOOL;                  // 保持中指示（bHold 电平镜像） [-] / Holding indicator
    eErrCode : E_DL_ShrErr;           // 信息码出口 / Info code outlet
    bError   : BOOL;                  // 故障标志（本件无故障级条件，恒 FALSE，契约位） [-] / Error flag, contract pin, always FALSE
END_VAR
VAR
    _abSnap  : ARRAY[0..7] OF BOOL;   // 锁存副本（唯一快照源，判定只读此副本） [-] / Latched snapshot, sole judgment source
    _uChg    : WORD;                  // 不一致位图内部锁存量（非恢复沿保持） [-] / Mismatch bitmap latch
    _bDiff   : BOOL;                  // 恢复沿存在不一致当拍量 [-] / Mismatch exists at resume
    i        : DINT;                  // 通道循环索引 / Channel loop index
    rtHold   : R_TRIG;                // 保持上升沿实例，段 0 无条件调用 / Hold rising-edge instance
    ftHold   : F_TRIG;                // 保持下降沿实例，段 0 无条件调用 / Hold falling-edge instance
END_VAR
VAR CONSTANT
    DL_SHR_NCHAN : DINT := 8;         // 通道定长 [路] / Fixed channel count
    DL_SHR_BIT0  : WORD := 1;         // bit0 基准掩码 [-] / Bit zero base mask
END_VAR

(* —— 段 0：沿实例无条件周期刷新（R6/R7） —— *)
rtHold(CLK := bHold);                 // 保持上升沿，每拍必调 / Hold rising edge, every scan
ftHold(CLK := bHold);                 // 保持下降沿，每拍必调 / Hold falling edge, every scan

(* —— 段 1：单拍量预清（_abSnap/_uChg 为锁存量不入清单，R107） —— *)
_bDiff := FALSE;                      // 不一致当拍量预清 / Mismatch preset

(* —— 段 2：保持上升沿 → 8 路拍照锁存 —— *)
IF rtHold.Q THEN
    FOR i := 0 TO (DL_SHR_NCHAN - 1) DO
        _abSnap[i] := abSignal[i];    // 逐通道快照锁存 / Per-channel snapshot latch
    END_FOR
END_IF

(* —— 段 3：恢复沿 → 锁存副本 vs 实时值逐通道一致性校验 —— *)
IF ftHold.Q THEN
    _uChg := 0;                       // 恢复沿重建位图（锁存量唯一写入点） / Rebuild bitmap at resume edge
    FOR i := 0 TO (DL_SHR_NCHAN - 1) DO
        IF _abSnap[i] <> abSignal[i] THEN
            _uChg := _uChg OR SHL(DL_SHR_BIT0, i);   // 不一致通道记位（i∈[0,7] 位宽内，结构性不越界） / Mark mismatch bit
            _bDiff := TRUE;           // 存在不一致 / Mismatch exists
        END_IF
    END_FOR
END_IF

(* —— 段 4：输出组合（保持期穿透闸：输出只取锁存副本） —— *)
FOR i := 0 TO (DL_SHR_NCHAN - 1) DO
    IF bHold THEN
        abOut[i] := _abSnap[i];       // 保持期：输出锁存副本（实时变化不穿透） / Held: output snapshot
    ELSE
        abOut[i] := abSignal[i];      // 恢复期：输出实时值 / Resumed: output live value
    END_IF
    abSnap[i] := _abSnap[i];          // 副本透读出口 / Snapshot readout outlet
END_FOR

(* —— 段 5：出口单点映射（名实双出口同源，R191） —— *)
bHolding := bHold;                    // 保持中指示（电平镜像） / Holding indicator
uChgMask := _uChg;                    // 位图出口（恢复沿外保持） / Bitmap outlet
IF _bDiff THEN
    eErrCode := E_DL_ShrErr.eResumeDiff;   // 信息级码（不置 bError） / Info code
ELSE
    eErrCode := E_DL_ShrErr.eOk;           // 一致或缺省 / Consistent or default
END_IF
bError := FALSE;                      // 本件无故障级条件（头注释声明，契约位恒 FALSE） / No fault-level condition

END_FUNCTION_BLOCK
